// ---- POUs/Tc3 Objects/Alarm/GVL_FB_Alarm_1.TcGVL
{attribute 'Tc2GvlVarNames'}
VAR_GLOBAL CONSTANT
	nALARM_MAX_NO			:INT := 63;			(* Maximal number of alarms *)
END_VAR

// ---- POUs/Tc3 Objects/Communication/TCPIP/GVL_TCPIP.TcGVL
{attribute 'qualified_only'}
VAR_GLOBAL CONSTANT
	BUFFER_SIZE						:UDINT := 1000;(* Max. internal fifo/receiver buffer size *)

	CLIENT_SEND_CYCLE_TIME			:TIME := T#1S;
	RECEIVE_POLLING_TIME			:TIME := T#100MS;
	RECEIVE_MESSAGE_MAX				:UINT := 10;

	(* Some project specific error codes *)
	ERROR_RECEIVE_TIMEOUT			:UDINT := 16#8101;(* Receive timeout *)
	ERROR_SENDFIFO_OVERFLOW			:UDINT := 16#8102;(* Send fifo overflow *)
	ERROR_RECFIFO_OVERFLOW			:UDINT := 16#8103;(* Receive fifo overflow *)
END_VAR

// ---- POUs/Tc3 Objects/ExternalHardware/Gefran/GVL_GFX4IR.TcGVL
{attribute 'qualified_only'}
VAR_GLOBAL CONSTANT
	nZONES_MAX_NO			:UINT := 4;			(* Amount of control zones *)
END_VAR

// ---- POUs/Tc3 Objects/File/CSV/GVL_CSV.TcGVL
VAR_GLOBAL CONSTANT
	MAX_CSV_ROWS 					:UDINT := 50;
	MAX_CSV_COLUMNS 				:UDINT := 50;
	MAX_CSV_FIELD_LENGTH			:UDINT := 100;
END_VAR

// ---- POUs/Tc3 Objects/File/TXT/GVL_FB_LoadFromFile_1.TcGVL
{attribute 'Tc2GvlVarNames'}
VAR_GLOBAL CONSTANT
	usnFileArrayMaxDimR					:USINT := 100;		(* 0..usnMaxDimR - Number of rows to read. *)
	usnFileArrayMaxDimC					:USINT := 4;  		(* 0..usnMaxDimC -  Number of columns to read. *)
END_VAR

// ---- POUs/Tc3 Objects/Logger/GVL_Logger.TcGVL
{attribute 'Tc2GvlVarNames'}
VAR_GLOBAL
	unLOG_INSTANCE_IDX				:UINT;
END_VAR
VAR_GLOBAL CONSTANT
	sLOG_FILE_PATH					:STRING := '\Hard Disk\Riex\Log\';			(* Login file path *)
	sLOG_FILE_SUFFIX					:STRING := 'log';							(* Suffix of loggin file *)
	unNUM_OF_LOG_VAR					:UINT := 4;								(* Number of logging variables *)
	unLOG_MAX_NO						:UINT := 1;
	unLOG_BEFOR_MAX_NO				:UINT := 10;
	unLOG_DURING_MAX_NO				:UINT := 250;
	unLOG_AFTER_MAX_NO				:UINT := 10;
END_VAR

// ---- POUs/Tc3 Objects/Traceability/GVL_Trace.TcGVL
{attribute 'Tc2GvlVarNames'}
VAR_GLOBAL CONSTANT
	MAX_TRACE_ROWS 					:UDINT := 1;
	MAX_TRACE_COLUMNS 				:UDINT := 30;
	MAX_TRACE_FIELD_LENGTH			:UDINT := 100;
END_VAR

// ---- POUs/MAIN.TcPOU
PROGRAM MAIN
VAR
	tonDelay			:TON;

	lrRight:LREAL;
	lrRight2:WORD;
	lrClamp2Pos:LREAL;
	lrActSawingAngle :LREAL;
END_VAR


Init();										(* Call Init *)
tonDelay(IN := TRUE, PT := t#3s);
Gr00Coordinator(bEnable := tonDelay.Q);			(* Call Program *)
Gr01Coordinator(bEnable := tonDelay.Q);			(* Call Program *)
Gr05Coordinator(bEnable := tonDelay.Q);			(* Call Program *)


lrActSawingAngle := (45 / 180 * PI);

lrClamp2Pos := F_AxisClamp2Pos(
					bEnable := TRUE,
					lrActClamp2Pos := Gr05Control.fbCylinderPos.lrActPosition,
					lrAngle := lrActSawingAngle,
					lrRadius := stgGr01HMI.stHMITOPLC.rPipeDiameter / 2.0,
					lrPipeClampWidth := lrgGr05PipeClampWidth,
					lrSawbandGuideWidth := lrgGr05SawbandGuideWidth
				);

lrRight := F_GetCylinderPos(		F_SetCylinderPos(SEL(stgGr05HMI.stHMITOPLC.bCylinderPosActive, Gr05Control.fbCylinderPos.lrActPosition, lrClamp2Pos),
																		lrgGr05CylinderPosOffset,
																		lrgGr05CylinderPosOriginShiftPos,
																		etgGr05CylinderPosDirection,
																		usngGr05CylinderPosCodingType),
														lrgGr05CylinderPosOffset,
														lrgGr05CylinderPosOriginShiftPos,
														etgGr05CylinderPosDirection,
														usngGr05CylinderPosCodingType)
									    + lrgGr05Clamp2Width ;



lrRight2 := F_SetCylinderPos(SEL(stgGr05HMI.stHMITOPLC.bCylinderPosActive, Gr05Control.fbCylinderPos.lrActPosition, lrClamp2Pos),
																		lrgGr05CylinderPosOffset,
																		lrgGr05CylinderPosOriginShiftPos,
																		etgGr05CylinderPosDirection,
																		usngGr05CylinderPosCodingType);

END_PROGRAM

// ---- POUs/Init.TcPOU
PROGRAM Init
VAR
	bFirstTime					:BOOL; 				(* False = first run / True = not first run *)
END_VAR
VAR PERSISTENT
	bFirstTimePersistent			:BOOL;				(* Persistente Daten initialisieren *)
END_VAR


IF NOT bFirstTime
THEN
	A_InitGr0000();
	A_InitGr0100();
	A_InitGr0200();
	A_InitGr0500();

	bFirstTime:= TRUE;
END_IF

IF NOT bFirstTimePersistent
THEN

	bFirstTimePersistent:= TRUE;
END_IF

ACTION A_InitGr0000:
;
END_ACTION

ACTION A_InitGr0100:
;
END_ACTION

ACTION A_InitGr0200:
;
END_ACTION

ACTION A_InitGr0500:
;
END_ACTION

END_PROGRAM

// ---- POUs/Machine/Group_0000 - General/Gr00Coordinator.TcPOU
PROGRAM Gr00Coordinator
VAR_INPUT
	(* Input variables / Eingang Variablen *)
	bEnable					:BOOL;						(* Enable Group00 *)
END_VAR
VAR
	(* Enummerations *)

	(* Variables *)

	(* References *)

	(* Interfaces *)

	(* Instances *)

END_VAR

IF NOT bEnable
THEN
	RETURN;
END_IF;

Gr00Persistent(bEnable := TRUE);			(* Call Program *)
Gr00Simulation(bEnable := TRUE);			(* Call Program *)
Gr00MachineMode(bEnable := TRUE);		(* Call Program *)
Gr00Control(bEnable := TRUE);				(* Call Program *)
Gr00HMI(bEnable := TRUE);				(* Call Program *)

END_PROGRAM

// ---- POUs/Machine/Group_0000 - General/Gr00Persistent/Gr00Persistent.TcPOU
PROGRAM Gr00Persistent
VAR_INPUT
	(* Input variables / Eingang Variablen *)
	bEnable					:BOOL;						(* Enable Gr00Persistent *)
END_VAR
VAR PERSISTENT
	(* Enummerations *)

	(* Variables *)
	rOverride							:REAL;						(* Override 0 - 100 % *)
	udnCounterTotal						:UDINT;						(* Total counter *)
	udnCounterUser						:UDINT;						(* User counter *)
	bProgramActive						:BOOL;						(* Program active *)

	arstSaveDiagSlaveInfo 				:ARRAY [0..dnDIAG_SLAVEINFO_SIZE] OF ST_SlaveStateInfo;
	arstSaveDiagSlaveInfoScanned			:ARRAY [0..dnDIAG_SLAVEINFO_SIZE] OF ST_SlaveStateInfoScanned;

	(* References *)

	(* Interfaces *)

	(* Instances *)
END_VAR
VAR
	(* Enummerations *)

	(* Variables *)
	bFirstTime							:BOOL;

	(* References *)

	(* Interfaces *)

	(* Instances *)

END_VAR

IF NOT bEnable
THEN
	bFirstTime := FALSE;
	RETURN;
END_IF;

IF NOT bFirstTime
THEN
	A_SetPerVar();

	bFirstTime := TRUE;
END_IF;

A_GetPerVar();

ACTION A_GetPerVar:

bgGr00WritePersistent := rOverride <> stgGr00HMI.stHMITOPLC.rOverride
					OR udnCounterTotal <> stgGr00HMI.stPLCTOHMI.udnCounterTotal
					OR udnCounterUser <> stgGr00HMI.stPLCTOHMI.udnCounterUser
					OR bProgramActive <> stgGr00HMI.stHMITOPLC.bProgramActive
					OR MEMCMP(ADR(arstSaveDiagSlaveInfo), ADR(SaveDiagSlaveInfo), SIZEOF(SaveDiagSlaveInfo)) <> 0
					OR MEMCMP(ADR(arstSaveDiagSlaveInfoScanned), ADR(SaveDiagSlaveInfoScanned), SIZEOF(SaveDiagSlaveInfoScanned)) <> 0;

rOverride := stgGr00HMI.stHMITOPLC.rOverride;
udnCounterTotal := stgGr00HMI.stPLCTOHMI.udnCounterTotal;
udnCounterUser := stgGr00HMI.stPLCTOHMI.udnCounterUser;
bProgramActive := stgGr00HMI.stHMITOPLC.bProgramActive;

MEMCPY(ADR(arstSaveDiagSlaveInfo), ADR(SaveDiagSlaveInfo), SIZEOF(SaveDiagSlaveInfo));
MEMCPY(ADR(arstSaveDiagSlaveInfoScanned), ADR(SaveDiagSlaveInfoScanned), SIZEOF(SaveDiagSlaveInfoScanned));
END_ACTION

ACTION A_SetPerVar:

stgGr00HMI.stHMITOPLC.rOverride := rOverride;
stgGr00HMI.stPLCTOHMI.udnCounterTotal := udnCounterTotal;
stgGr00HMI.stPLCTOHMI.udnCounterUser := udnCounterUser;
stgGr00HMI.stHMITOPLC.bProgramActive := bProgramActive;

MEMCPY(ADR(SaveDiagSlaveInfo), ADR(arstSaveDiagSlaveInfo), SIZEOF(arstSaveDiagSlaveInfo));
MEMCPY(ADR(SaveDiagSlaveInfoScanned), ADR(arstSaveDiagSlaveInfoScanned), SIZEOF(arstSaveDiagSlaveInfoScanned));
END_ACTION

END_PROGRAM

// ---- POUs/Machine/Group_0000 - General/Gr00Simulation/Gr00Simulation.TcPOU
PROGRAM Gr00Simulation
VAR_INPUT
	(* Input variables / Eingang Variablen *)
	bEnable								:BOOL;						(* Enable Gr05Persistent *)
END_VAR
VAR
	(* Enummerations *)

	(* Variables *)

	(* References *)

	(* Interfaces *)

	(* Instances *)

END_VAR

IF NOT bEnable
THEN

	RETURN;
END_IF;

A_ForceInput();

ACTION A_ForceInput:


GVL_Gr00IO.binGr00AirPressureOK := TRUE;
GVL_Gr00IO.binGr00LightCurtainOK := TRUE;
GVL_Gr00IO.arbinGr00PowerSupplyOn[2] := TRUE;
GVL_Gr00IO.arbinGr00PowerSupplyOn[3] := TRUE;
GVL_Gr00IO.arbinGr00PowerSupplyOn[4] := TRUE;
GVL_Gr00IO.arbinGr00PowerSupplyOn[5] := TRUE;
GVL_Gr00IO.arbinGr00DoorsClosed[1] := TRUE;
GVL_Gr00IO.arbinGr00DoorsClosed[2] := TRUE;
GVL_Gr00IO.arbinGr00DoorsClosed[3] := TRUE;
GVL_Gr00IO.arbinGr00DoorsClosed[4] := TRUE;
GVL_Gr00IO.arbinGr00DoorsClosed[5] := TRUE;
GVL_Gr00IO.binGr00AllDoorsClosed := GVL_Gr00IO.arbinGr00DoorsClosed[1]
								AND GVL_Gr00IO.arbinGr00DoorsClosed[2]
								AND GVL_Gr00IO.arbinGr00DoorsClosed[3]
								AND GVL_Gr00IO.arbinGr00DoorsClosed[4]
								AND GVL_Gr00IO.arbinGr00DoorsClosed[5];

GVL_Gr00IO.binGr00AllDoorsLocked := TRUE;
GVL_Gr00IO.binGr00TempOK := TRUE;


// only for simulation
// GVL_Gr00IO.binNoEmergencyStop := TRUE;
// GVL_Gr00IO.binMoveRelease := TRUE;
// GVL_Gr00IO.binMoveReleaseSB := TRUE;
END_ACTION

END_PROGRAM

// ---- POUs/Machine/Group_0000 - General/Gr00MachineMode/Gr00MachineMode.TcPOU
PROGRAM Gr00MachineMode
VAR_INPUT
	(* Input variables / Eingang Variablen *)
	bEnable					:BOOL;						(* Enable Gr00MachineMode *)
END_VAR
VAR
	(* Enummerations *)

	(* Variables *)

	(* References *)

	(* Interfaces *)

	(* Instances *)

END_VAR

IF NOT bEnable
THEN
	RETURN;
END_IF;

Gr00Auto(bEnable := TRUE);			(* Call Program *)
Gr00Home(bEnable := TRUE);			(* Call Program *)
Gr00Manual(bEnable := TRUE);			(* Call Program *)

END_PROGRAM

// ---- POUs/Machine/Group_0000 - General/Gr00MachineMode/Gr00Auto/Gr00Auto.TcPOU
PROGRAM Gr00Auto
VAR_INPUT
	(* Input variables / Eingang Variablen *)
	bEnable					:BOOL;						(* Enable Gr00Auto *)
	bExecute				:BOOL;						(* Auto execute *)

	(* Instances *)
	fbInit						:FB_Gr00AutoInit;
	fbProcedure				:FB_Gr00AutoProcedure;
END_VAR
VAR
	(* Enummerations *)

	(* Variables *)

	(* References *)

	(* Interfaces *)

	(* Instances *)
	rtExecute					:R_TRIG;

	fbAlarm					:FB_Gr00AutoAlarm;
END_VAR
VAR CONSTANT
	nFatalErrorMaxIdx				:INT := 0;						(* Maximal index of  using alarms *)
	nErrorMaxIdx					:INT := 0;						(* Maximal index of  using alarms *)
	nWarningMaxIdx				:INT := 0;						(* Maximal index of  using alarms *)
	nMessageMaxIdx				:INT := 0;						(* Maximal index of  using alarms *)
	nHintMaxIdx					:INT := 0;						(* Maximal index of  using alarms *)

	dnFatalErrorBaseIdentNo		:DINT := 02000;				(* Fatal error identification number *)
	dnErrorBaseIdentNo			:DINT := 02100;				(* Error identification number *)
	dnWarningBaseIdentNo		:DINT := 02200;				(* Warning identification number *)
	dnMessageBaseIdentNo		:DINT := 02300;				(* Message identification number *)
	dnHintBaseIdentNo			:DINT := 02400;				(* Hint identification number *)
END_VAR

IF NOT bEnable
THEN
    RETURN;
END_IF;

(* Check auto execute *)
bExecute := bgGr00ModeAutomatic
		      AND NOT fbInit.bFirstTime;

rtExecute(CLK := bExecute);

IF rtExecute.Q
THEN
	A_Init();
END_IF;

A_Procedure();
A_Alarm();

ACTION A_Alarm:

(* Collect and execute input alarms *)
fbAlarm.stAlarmIn.arbError[0].bActive := FALSE;
fbAlarm.stAlarmIn.arbError[0].dnCode := dnErrorBaseIdentNo + 0;

fbAlarm(
	etMachineMode := etgGr00MachineMode,
	etMachineState := etgGr00MachineState,
	bNoEStop := bgGr00NoEmergencyStop,
	bConfirmAlarm := bgGr00ConfirmAlarm,
	dtDateTime := stgGr00DateTime.dtDateTime,
	nFatalErrorMaxIdx := nFatalErrorMaxIdx,
	nErrorMaxIdx := nErrorMaxIdx,
	nWarningMaxIdx := nWarningMaxIdx,
	nMessageMaxIdx := nMessageMaxIdx,
	nHintMaxIdx := nHintMaxIdx,
	bMoveInterrupted := bgGr00MoveInterrupted,
	bHomeCompleted := bgGr00HomeCompleted,
	stAlarmOut => stgGr00Alarm.stAuto
);
END_ACTION

ACTION A_Init:

(* Initializing variables *)
fbInit();
END_ACTION

ACTION A_Procedure:

(* Execute auto procedure *)
fbProcedure(
	bEnable := fbInit.bFirstTime,
	bExecute := etgGr00MachineState = ET_MachineState_eAutoExe
	             	       OR etgGr00MachineState = ET_MachineState_eAutoSteppingExe,
	bInterrupt := FALSE,
	bReleaseNextStep := etgGr00MachineState = ET_MachineState_eAutoExe
	             	       		       OR etgGr00MachineState = ET_MachineState_eAutoSteppingExe,
	bDone => bgGr00AutoCompleted,
	bInterrupted => bgGr00MoveInterrupted
);
END_ACTION

END_PROGRAM

// ---- POUs/Machine/Group_0000 - General/Gr00MachineMode/Gr00Home/Gr00Home.TcPOU
PROGRAM Gr00Home
VAR_INPUT
	(* Input variables / Eingang Variablen *)
	bEnable					:BOOL;						(* Enable Gr00Home *)
	bExecute				:BOOL;						(* Home execute *)

	(* Instances *)
	fbInit						:FB_Gr00HomeInit;
	fbProcedure				:FB_Gr00HomeProcedure;
END_VAR
VAR
	(* Enummerations *)

	(* Variables *)

	(* References *)

	(* Interfaces *)

	(* Instances *)
	rtExecute					:R_TRIG;

	fbAlarm					:FB_Gr00HomeAlarm;

END_VAR
VAR CONSTANT
	nFatalErrorMaxIdx				:INT := 0;						(* Maximal index of  using alarms *)
	nErrorMaxIdx					:INT := 0;						(* Maximal index of  using alarms *)
	nWarningMaxIdx				:INT := 0;						(* Maximal index of  using alarms *)
	nMessageMaxIdx				:INT := 0;						(* Maximal index of  using alarms *)
	nHintMaxIdx					:INT := 0;						(* Maximal index of  using alarms *)

	dnFatalErrorBaseIdentNo		:DINT := 03000;				(* Fatal error identification number *)
	dnErrorBaseIdentNo			:DINT := 03100;				(* Error identification number *)
	dnWarningBaseIdentNo		:DINT := 03200;				(* Warning identification number *)
	dnMessageBaseIdentNo		:DINT := 03300;				(* Message identification number *)
	dnHintBaseIdentNo			:DINT := 03400;				(* Hint identification number *)
END_VAR

IF NOT bEnable
THEN
	RETURN;
END_IF;

(* Check home execute *)
bExecute := etgGr00MachineState = ET_MachineState_eHomeRefExe
		      OR etgGr00MachineState = ET_MachineState_eHomeExe;

rtExecute(CLK := bExecute);                   

IF rtExecute.Q
THEN
	fbInit.bFirstTime := FALSE;
	A_Init();
END_IF;

A_Procedure();
A_Alarm();

ACTION A_Alarm:

(* Collect and execute input alarms *)
fbAlarm.stAlarmIn.arbError[0].bActive := fbProcedure.bErrorByProgramVerification;
fbAlarm.stAlarmIn.arbError[0].dnCode := dnErrorBaseIdentNo + 0;

fbAlarm(
	etMachineMode := etgGr00MachineMode,
	etMachineState := etgGr00MachineState,
	bNoEStop := bgGr00NoEmergencyStop,
	bConfirmAlarm := bgGr00ConfirmAlarm,
	dtDateTime := stgGr00DateTime.dtDateTime,
	nFatalErrorMaxIdx := nFatalErrorMaxIdx,
	nErrorMaxIdx := nErrorMaxIdx,
	nWarningMaxIdx := nWarningMaxIdx,
	nMessageMaxIdx := nMessageMaxIdx,
	nHintMaxIdx := nHintMaxIdx,
	bMoveInterrupted := bgGr00MoveInterrupted,
	bHomeCompleted := bgGr00HomeCompleted,
	stAlarmOut => stgGr00Alarm.stHome
);
END_ACTION

ACTION A_Init:

(* Initializing variables *)
fbInit();
END_ACTION

ACTION A_Procedure:

(* Execute home procedure *)
fbProcedure(
	bEnable := etgGr00MachineMode = ET_MachineMode_eHome,
	bExecute := rtExecute.Q,
	bReleaseNextStep := etgGr00MachineState = ET_MachineState_eHomeRefExe
		      	     		      OR etgGr00MachineState = ET_MachineState_eHomeExe
);
END_ACTION

END_PROGRAM

// ---- POUs/Machine/Group_0000 - General/Gr00MachineMode/Gr00Manual/Gr00Manual.TcPOU
PROGRAM Gr00Manual
VAR_INPUT
	(* Input variables / Eingang Variablen *)
	bEnable					:BOOL;						(* Enable Gr00Manual *)
	bExecute				:BOOL;						(* Manual execute *)

	(* Instances *)
	fbInit						:FB_Gr00ManualInit;
	fbProcedure				:FB_Gr00ManualProcedure;
END_VAR
VAR
	(* Enummerations *)

	(* Variables *)

	(* References *)

	(* Interfaces *)

	(* Instances *)
	rtExecute					:R_TRIG;

	fbAlarm					:FB_Gr00ManualAlarm;
END_VAR
VAR CONSTANT
	nFatalErrorMaxIdx				:INT := 0;						(* Maximal index of  using alarms *)
	nErrorMaxIdx					:INT := 0;						(* Maximal index of  using alarms *)
	nWarningMaxIdx				:INT := 0;						(* Maximal index of  using alarms *)
	nMessageMaxIdx				:INT := 0;						(* Maximal index of  using alarms *)
	nHintMaxIdx					:INT := 0;						(* Maximal index of  using alarms *)

	dnFatalErrorBaseIdentNo		:DINT := 04000;				(* Fatal error identification number *)
	dnErrorBaseIdentNo			:DINT := 04100;				(* Error identification number *)
	dnWarningBaseIdentNo		:DINT := 04200;				(* Warning identification number *)
	dnMessageBaseIdentNo		:DINT := 04300;				(* Message identification number *)
	dnHintBaseIdentNo			:DINT := 04400;				(* Hint identification number *)
END_VAR

IF NOT bEnable
THEN
	RETURN;
END_IF;

(* Check manual execute *)
bExecute := etgGr00MachineMode = ET_MachineMode_eManual;

rtExecute(CLK := bExecute);

IF rtExecute.Q
THEN
	fbInit.bFirstTime := FALSE;
	A_Init();
END_IF;

A_Procedure();
A_Alarm();

ACTION A_Alarm:

(* Collect and execute input alarms *)
fbAlarm.stAlarmIn.arbError[0].bActive := FALSE;
fbAlarm.stAlarmIn.arbError[0].dnCode := dnErrorBaseIdentNo + 0;

fbAlarm(
	etMachineMode := etgGr00MachineMode,
	etMachineState := etgGr00MachineState,
	bNoEStop := bgGr00NoEmergencyStop,
	bConfirmAlarm := bgGr00ConfirmAlarm,
	dtDateTime := stgGr00DateTime.dtDateTime,
	nFatalErrorMaxIdx := nFatalErrorMaxIdx,
	nErrorMaxIdx := nErrorMaxIdx,
	nWarningMaxIdx := nWarningMaxIdx,
	nMessageMaxIdx := nMessageMaxIdx,
	nHintMaxIdx := nHintMaxIdx,
	bHomeCompleted := bgGr00HomeCompleted,
	stAlarmOut => stgGr00Alarm.stManual
);
END_ACTION

ACTION A_Init:

(* Initializing variables *)
fbInit();
END_ACTION

ACTION A_Procedure:

(* Execute manual procedure *)
fbProcedure(
	bEnable := etgGr00MachineMode = ET_MachineMode_eManual,
	bExecute := rtExecute.Q,
	bReleaseNextStep := etgGr00MachineMode = ET_MachineMode_eManual
);
END_ACTION

END_PROGRAM

// ---- POUs/Machine/Group_0000 - General/Gr00Control/Gr00Control.TcPOU
PROGRAM Gr00Control
VAR_INPUT
	(* Input variables / Eingang Variablen *)
	bEnable					:BOOL;						(* Enable Gr00Control *)

	fbProgram				:FB_Gr00Program;
END_VAR
VAR
	(* Enummerations *)

	(* Variables *)

	(* References *)

	(* Interfaces *)

	(* Instances *)
	fbAlarm					:FB_Gr00Alarm;
	fbSafety					:FB_Gr00Safety;
	fbSignals				:FB_Gr00Signals;
	fbUtility					:FB_Gr00Utility;
	fbPeriphery				:FB_Gr00Periphery;

	ftClampsChecked			:F_TRIG;
	tonClampsChecked		:TON;
	fbMachineStandstill		:FB_SignalHandlingDelay;

	fbStartHMI				:NT_StartProcess;
	tonStartHmi				:TON;

END_VAR
VAR CONSTANT
	nFatalErrorMaxIdx				:INT := 1;						(* Maximal index of  using alarms *)
	nErrorMaxIdx					:INT := 12;					(* Maximal index of  using alarms *)
	nWarningMaxIdx				:INT := 0;						(* Maximal index of  using alarms *)
	nMessageMaxIdx				:INT := 4;						(* Maximal index of  using alarms *)
	nHintMaxIdx					:INT := 0;						(* Maximal index of  using alarms *)

	dnFatalErrorBaseIdentNo		:DINT := 01000;				(* Fatal error identification number *)
	dnErrorBaseIdentNo			:DINT := 01100;				(* Error identification number *)
	dnWarningBaseIdentNo		:DINT := 01200;				(* Warning identification number *)
	dnMessageBaseIdentNo		:DINT := 01300;				(* Message identification number *)
	dnHintBaseIdentNo			:DINT := 01400;				(* Hint identification number *)
END_VAR

IF NOT bEnable
THEN
	RETURN;
END_IF;

A_Periphery();
A_Utility();
A_Program();
A_Safety();
A_Signals();
A_Alarm();
A_HMI();

ACTION A_Alarm:

(* Collect and execute input alarms *)
fbAlarm.stAlarmIn.arbFatalError[0].bActive := fbSafety.fbNoEmergencyStop.bError;
fbAlarm.stAlarmIn.arbFatalError[0].dnCode := dnFatalErrorBaseIdentNo + 0;

fbAlarm.stAlarmIn.arbError[0].bActive := NOT binGr00LightCurtainOK
                                                		      AND (Gr01Home.fbProcedure.bBusy
                                                      				OR Gr01Auto.fbProcedure.bBusy);
fbAlarm.stAlarmIn.arbError[0].dnCode := dnErrorBaseIdentNo + 0;

fbAlarm.stAlarmIn.arbError[1].bActive := fbSafety.fbAirPressure.bError;
fbAlarm.stAlarmIn.arbError[1].dnCode := dnErrorBaseIdentNo + 1;

fbAlarm.stAlarmIn.arbError[2].bActive := FALSE;
fbAlarm.stAlarmIn.arbError[2].dnCode := dnErrorBaseIdentNo + 2;

fbAlarm.stAlarmIn.arbError[4].bActive := NOT fbSafety.bFieldbusMasterOK AND fbSafety.fbFieldbus.bInit;
fbAlarm.stAlarmIn.arbError[4].dnCode := dnErrorBaseIdentNo + 4;

fbAlarm.stAlarmIn.arbError[5].bActive := fbSafety.bFieldbusBrake;
fbAlarm.stAlarmIn.arbError[5].dnCode := dnErrorBaseIdentNo + 5;

fbAlarm.stAlarmIn.arbError[6].bActive := fbSafety.fbTemperatur.bError;
fbAlarm.stAlarmIn.arbError[6].dnCode := dnErrorBaseIdentNo + 6;

fbAlarm.stAlarmIn.arbError[7].bActive := NOT fbSafety.arbPowerSupplyOn[1];
fbAlarm.stAlarmIn.arbError[7].dnCode := dnErrorBaseIdentNo + 7;

fbAlarm.stAlarmIn.arbError[8].bActive :=NOT fbSafety.arbPowerSupplyOn[2];
fbAlarm.stAlarmIn.arbError[8].dnCode := dnErrorBaseIdentNo + 8;

fbAlarm.stAlarmIn.arbError[9].bActive := NOT fbSafety.arbPowerSupplyOn[3];
fbAlarm.stAlarmIn.arbError[9].dnCode := dnErrorBaseIdentNo + 9;

fbAlarm.stAlarmIn.arbError[10].bActive := FALSE(*SystemInfo.bootDataFlags.5*);
fbAlarm.stAlarmIn.arbError[10].dnCode := dnErrorBaseIdentNo + 10;

fbAlarm.stAlarmIn.arbError[11].bActive := fbProgram.fbRead.bError
								      AND  fbProgram.fbRead.udnErrorNo <> 31;
fbAlarm.stAlarmIn.arbError[11].dnCode := dnErrorBaseIdentNo + 11;

fbAlarm.stAlarmIn.arbError[12].bActive := fbProgram.fbRead.bError
								      AND  fbProgram.fbRead.udnErrorNo = 31;
fbAlarm.stAlarmIn.arbError[12].dnCode := dnErrorBaseIdentNo + 12;

fbAlarm.stAlarmIn.arbWarning[0].bActive := fbSafety.fbTemperatur.bWarning;
fbAlarm.stAlarmIn.arbWarning[0].dnCode := dnWarningBaseIdentNo + 0;

fbAlarm.stAlarmIn.arbWarning[1].bActive := NOT GVL_Gr00IO.binGr00Luetze_F1;
fbAlarm.stAlarmIn.arbWarning[1].dnCode := dnWarningBaseIdentNo + 1;

fbAlarm.stAlarmIn.arbWarning[2].bActive := NOT GVL_Gr00IO.binGr00Luetze_F2;
fbAlarm.stAlarmIn.arbWarning[2].dnCode := dnWarningBaseIdentNo + 2;

fbAlarm.stAlarmIn.arbWarning[3].bActive := NOT GVL_Gr00IO.binGr00Luetze_F3;
fbAlarm.stAlarmIn.arbWarning[3].dnCode := dnWarningBaseIdentNo + 3;

fbAlarm.stAlarmIn.arbWarning[4].bActive := NOT GVL_Gr00IO.binGr00PS6A24Warning_1;
fbAlarm.stAlarmIn.arbWarning[4].dnCode := dnWarningBaseIdentNo + 4;

fbAlarm.stAlarmIn.arbWarning[5].bActive := NOT GVL_Gr00IO.binGr00PS6A24Warning_2;
fbAlarm.stAlarmIn.arbWarning[5].dnCode := dnWarningBaseIdentNo + 5;

fbAlarm.stAlarmIn.arbWarning[6].bActive := NOT GVL_Gr00IO.binGr00PS6A24Ready;
fbAlarm.stAlarmIn.arbWarning[6].dnCode := dnWarningBaseIdentNo + 6;

fbAlarm.stAlarmIn.arbMessage[0].bActive := fbSafety.fbAirPressure.udnMessageNo = 1;
fbAlarm.stAlarmIn.arbMessage[0].dnCode := dnMessageBaseIdentNo + 0;

fbAlarm.stAlarmIn.arbMessage[1].bActive := stgGr00HMI.stHMITOPLC.bSafetyInterlockOff;
fbAlarm.stAlarmIn.arbMessage[1].dnCode := dnMessageBaseIdentNo + 1;

fbAlarm.stAlarmIn.arbMessage[2].bActive := NOT binGr00LightCurtainOK
                                            				      AND NOT fbAlarm.stAlarmIn.arbError[0].bActive
                                            				      AND NOT stgGr00Alarm.stControl.arbError[0].bActive;
fbAlarm.stAlarmIn.arbMessage[2].dnCode := dnMessageBaseIdentNo + 2;

fbAlarm.stAlarmIn.arbMessage[4].bActive := NOT binGr00AllDoorsClosed;
fbAlarm.stAlarmIn.arbMessage[4].dnCode := dnMessageBaseIdentNo + 4;

(* Execute utility *)
fbAlarm(
	etMachineMode := etgGr00MachineMode,
	etMachineState := etgGr00MachineState,
	bNoEStop := bgGr00NoEmergencyStop,
	bConfirmAlarm := bgGr00ConfirmAlarm,
	dtDateTime := stgGr00DateTime.dtDateTime,
	nFatalErrorMaxIdx := nFatalErrorMaxIdx,
	nErrorMaxIdx := nErrorMaxIdx,
	nWarningMaxIdx := nWarningMaxIdx,
	nMessageMaxIdx := nMessageMaxIdx,
	nHintMaxIdx := nHintMaxIdx,
	bMoveInterrupted := bgGr00MoveInterrupted,
	bHomeCompleted := bgGr00HomeCompleted,
	stAlarmOut => stgGr00Alarm.stControl
);
END_ACTION

ACTION A_HMI:
(*Starting the HMI*)

tonStartHmi(IN:=TRUE, PT:= T#2s);

fbStartHMI(
		PATHSTR   := 'C:\Riex\HMI\App.exe',
    		DIRNAME   :='C:\Riex\HMI\',
    		START     := tonStartHmi.Q,
		TMOUT     := T#5s
		);
END_ACTION

ACTION A_Periphery:

(* Periphery *)
fbPeriphery(
	bEnable := TRUE,
	Periphery := Periphery
);
END_ACTION

ACTION A_Program:

(* Execute program *)
fbProgram(
	sPath := sgGr00PrgPath,
	sName := sgGr00PrgName,
	sSuffix := sgGr00PrgSuffix
);
END_ACTION

ACTION A_Safety:

bgGr00DoorsUnlockRelease := bgGr00ModeManual
						        OR
							(bgGr00ModeHome
							 AND NOT bgGr00MachineRunning)
						        OR
							(bgGr00ModeAutomatic
							 AND NOT bgGr00MachineRunning);

(* Execute safety *)
fbSafety(
	etMachineMode := etgGr00MachineMode,
	etMachineState := etgGr00MachineState,
	bNoEStop := binGr00NoEmergencyStop,
	bConfirmEStop := FALSE,
	bMachineRunning := bgGr00MachineRunning,
	arbPowerSupplyOn := arbinGr00PowerSupplyOn,
	bLightCurtain := binGr00LightCurtainOK,
	bConfirmLightCurtain := (bgGr00ConfirmAlarm
						OR etgGr00MachineMode = ET_MachineMode_eManual
						OR etgGr00MachineMode = ET_MachineMode_eHome
						OR etgGr00MachineMode = ET_MachineMode_eAutomatic
						OR stgGr00HMI.stHMITOPLC.bSafetyInterlockOff)
						AND NOT stgGr00Alarm.stControl.arbError[0].bActive,
	bAirPressure := binGr00AirPressureOK,
	arbDoorsClosed := arbinGr00DoorsClosed,
	bDoorsClosed := binGr00AllDoorsClosed,
	bDoorsLocked := binGr00AllDoorsLocked,
	bTemperatur := binGr00TempOK,
	stFieldbusStatus := stinGr00FieldbusStatus,
	tFieldbusMasterStartUp := tgGr00FieldbusMasterStartUp,
	tPowerSupplyOn := tgGr00PowerSupplyOn,
	tPowerSupplyOff := tgGr00PowerSupplyOff,
	tAirPressureOnDelay := tgGr00AirPressureOnDelay,
	tAirPresentDelay := tgGr00AirPressureDelay,
	tAirPressureBuildUp := tgGr00AirPressureBuildUp,
	tLightCurtainDelay := tgGr00LightCurtainDelay,
	tAdsTimeOut := DEFAULT_ADS_TIMEOUT,
	bNoEmergencyStop => bgGr00NoEmergencyStop,
	bAirPressureOK => bgGr00AirPressureOK,
	bAirPressureOn => boutGr00AirPressureOn,
	bPowerSupplyOk => bgGr00PowerSupplyOk,
	bLightCurtainOK => bgGr00LightCurtainOK,
	bConfirmedLightCurtain => boutGr00ConfLightCurtain,
	bAllDoorsLock => boutGr00AllDoorsLock,
	bAllDoorsClosed => bgGr00AllDoorsClosed,
	bAllDoorsClosedLocked => bgGr00AllDoorsClosedLocked
);
END_ACTION

ACTION A_Signals:

(* Collect and execute input signals *)
fbSignals.stAlarm.bFatalError := stgGr00Alarm.stControl.bFatalError OR stgGr00Alarm.stManual.bFatalError OR stgGr00Alarm.stHome.bFatalError OR stgGr00Alarm.stAuto.bFatalError
							OR stgGr01Alarm.stControl.bFatalError OR stgGr01Alarm.stManual.bFatalError OR stgGr01Alarm.stHome.bFatalError OR stgGr01Alarm.stAuto.bFatalError
							OR stgGr02Alarm.stControl.bFatalError OR stgGr02Alarm.stManual.bFatalError OR stgGr02Alarm.stHome.bFatalError OR stgGr02Alarm.stAuto.bFatalError
							OR stgGr05Alarm.stControl.bFatalError OR stgGr05Alarm.stManual.bFatalError OR stgGr05Alarm.stHome.bFatalError OR stgGr05Alarm.stAuto.bFatalError;
fbSignals.stAlarm.bError := stgGr00Alarm.stControl.bError OR stgGr00Alarm.stManual.bError OR stgGr00Alarm.stHome.bError OR stgGr00Alarm.stAuto.bError
						OR stgGr01Alarm.stControl.bError OR stgGr01Alarm.stManual.bError OR stgGr01Alarm.stHome.bError OR stgGr01Alarm.stAuto.bError
						OR stgGr02Alarm.stControl.bError OR stgGr02Alarm.stManual.bError OR stgGr02Alarm.stHome.bError OR stgGr02Alarm.stAuto.bError
						OR stgGr05Alarm.stControl.bError OR stgGr05Alarm.stManual.bError OR stgGr05Alarm.stHome.bError OR stgGr05Alarm.stAuto.bError;
fbSignals.stAlarm.bWarning := stgGr00Alarm.stControl.bWarning OR stgGr00Alarm.stManual.bWarning OR stgGr00Alarm.stHome.bWarning OR stgGr00Alarm.stAuto.bWarning
		        					OR stgGr01Alarm.stControl.bWarning OR stgGr01Alarm.stManual.bWarning OR stgGr01Alarm.stHome.bWarning OR stgGr01Alarm.stAuto.bWarning
		        					OR stgGr02Alarm.stControl.bWarning OR stgGr02Alarm.stManual.bWarning OR stgGr02Alarm.stHome.bWarning OR stgGr02Alarm.stAuto.bWarning
		        					OR stgGr05Alarm.stControl.bWarning OR stgGr05Alarm.stManual.bWarning OR stgGr05Alarm.stHome.bWarning OR stgGr05Alarm.stAuto.bWarning;
fbSignals.stAlarm.bMessage := stgGr00Alarm.stControl.bMessage OR stgGr00Alarm.stManual.bMessage OR stgGr00Alarm.stHome.bMessage OR stgGr00Alarm.stAuto.bMessage
		        					OR stgGr01Alarm.stControl.bMessage OR stgGr01Alarm.stManual.bMessage OR stgGr01Alarm.stHome.bMessage OR stgGr01Alarm.stAuto.bMessage
		        					OR stgGr02Alarm.stControl.bMessage OR stgGr02Alarm.stManual.bMessage OR stgGr02Alarm.stHome.bMessage OR stgGr02Alarm.stAuto.bMessage
		        					OR stgGr05Alarm.stControl.bMessage OR stgGr05Alarm.stManual.bMessage OR stgGr05Alarm.stHome.bMessage OR stgGr05Alarm.stAuto.bMessage;
fbSignals.stAlarm.bHint := stgGr00Alarm.stControl.bHint OR stgGr00Alarm.stManual.bHint OR stgGr00Alarm.stHome.bHint OR stgGr00Alarm.stAuto.bHint
	       					OR stgGr01Alarm.stControl.bHint OR stgGr01Alarm.stManual.bHint OR stgGr01Alarm.stHome.bHint OR stgGr01Alarm.stAuto.bHint
	       					OR stgGr02Alarm.stControl.bHint OR stgGr02Alarm.stManual.bHint OR stgGr02Alarm.stHome.bHint OR stgGr02Alarm.stAuto.bHint
	       					OR stgGr05Alarm.stControl.bHint OR stgGr05Alarm.stManual.bHint OR stgGr05Alarm.stHome.bHint OR stgGr05Alarm.stAuto.bHint;

(* Execute signals *)
fbSignals(
	etMachineMode := etgGr00MachineMode,
	etMachineState := etgGr00MachineState,
	bMachineRunning := bgGr00MachineRunning,
	stBlinker => stgGr00Blinker,
	bBulbBtnStart => boutGr00BulbBtnStart,
	bBulbBtnStop => boutGr00BulbBtnStop,
	bBulbBtnHome => boutGr00BulbBtnHome,
	bBulbGreen => boutGr00BulbGreen,
	bBulbRed => boutGr00BulbRed,
	bBulbYellow => boutGr00BulbYellow,
	bHorn => boutGr00Horn
);

(* Signal button bulb "reset" / Signallampe "Reset" *)
boutGr00BulbBtnReset := binGr00NoEmergencyStop OR stgGr00Blinker.Q1;
END_ACTION

ACTION A_Utility:

(* Execute utility *)
fbUtility(
	bSignalStart := binGr00PushBtnStart OR stgGr00HMI.stHMITOPLC.bBtnStart,
	bSignalStop :=NOT binGr00PushBtnStop OR stgGr00HMI.stHMITOPLC.bBtnStop,
	bSignalAbort := fbSignals.stAlarm.bFatalError
				     OR fbSignals.stAlarm.bError,
	bSignalHome := binGr00PushBtnHome,
	bSignalReference := binGr00PushBtnRef OR stgGr00HMI.stHMITOPLC.bBtnForceRef,
	bSignalReset := binGr00PushBtnReset OR stgGr00HMI.stHMITOPLC.bBtnReset,
	bSignalMachinePurge := stgGr00HMI.stHMITOPLC.bBtnMachinePurge,
	bAutoStartRelease := binGr01SawbandRelease
					       AND bgGr05PipeEndPresent
					       AND (stgGr05HMI.stHMITOPLC.bCylinderPosActive
							  OR stgGr05HMI.stPLCTOHMI.arlrAxisClampActPos[2] < ABS(99999.0))
					       AND NOT stgGr05Alarm.stAuto.arbWarning[0].bActive,
	bHomeStartRelease := (stgGr05HMI.stHMITOPLC.bCylinderPosActive
							  OR stgGr05HMI.stPLCTOHMI.arlrAxisClampActPos[2] < ABS(99999.0)),
	bAutoToHome := NOT stgGr05Alarm.stAuto.arbWarning[0].bActive,
	bHomeCompleted := bgGr00HomeCompleted
					     AND bgGr01HomeCompleted
					     AND bgGr02HomeCompleted
					     AND bgGr05HomeCompleted,
	bAutoCompleted := bgGr00AutoCompleted
					  AND bgGr01AutoCompleted
					  AND bgGr02AutoCompleted
					  AND bgGr05AutoCompleted,
	bAllDoorsClosed := binGr00AllDoorsClosed,
	bAllDoorsLocked := bgGr00AllDoorsClosedLocked,
	bLightCurtainOk := bgGr00LightCurtainOK,
	etMachineModeReq := stgGr00HMI.stHMITOPLC.etMachineMode,
	bExeCounter := bgGr00AutoCompleted
					  AND bgGr01AutoCompleted
					  AND bgGr02AutoCompleted
					  AND bgGr05AutoCompleted,
	bResetCounterUser := stgGr00HMI.stHMITOPLC.bResetCounterUser,
	bStartTime := Gr01Control.fbUtility.arbStartProcess[1]
				OR Gr01Control.fbUtility.arbStartProcess[2]
				OR Gr01Control.fbUtility.arbStartProcess[3],
	bStopTime := bgGr01AutoCompleted
				OR Gr01Control.fbUtility.arbStopProcess[1]
				OR Gr01Control.fbUtility.arbStopProcess[2]
				OR Gr01Control.fbUtility.arbStopProcess[3],
	bLifetimeOn := TRUE,
	bResetLifetimeAll := FALSE,
	sLifetimeFilePath := sgGr00MachineLifetimeFilePath,
	sLifetimeFileName := sgGr00MachineLifetimeFileName,
	bWritePersistent :=  bgGr00WritePersistent
					  OR  bgGr01WritePersistent
					  OR  bgGr02WritePersistent
					  OR  bgGr05WritePersistent,
	bDownTraceDataExe := FALSE,
	rGlobalOverride := stgGr00HMI.stHMITOPLC.rOverride,
	udnCounterTotal := stgGr00HMI.stPLCTOHMI.udnCounterTotal,
	udnCounterUser := stgGr00HMI.stPLCTOHMI.udnCounterUser,
	tAdsTimeOut := DEFAULT_ADS_TIMEOUT,
	etMachineMode => etgGr00MachineMode,
	etMachineState => etgGr00MachineState,
	bModeAutomatic => bgGr00ModeAutomatic,
	bModeHome => bgGr00ModeHome,
	bModeManual => bgGr00ModeManual,
	bMachineRunning => bgGr00MachineRunning,
	bMachineStandstill => bgGr00MachineStandstill,
	bMachinePurge => bgGr00MachinePurge,
	bConfirmAlarm => bgGr00ConfirmAlarm,
	rActOverride => rgGr00Override,
	lrLifetimeAll => stgGr00HMI.stPLCTOHMI.lrMachineLifetime,
	lrLifetimeAfterTrunOn => stgGr00HMI.stPLCTOHMI.lrMachineLifetimeAfterTurnOn,
	lrActCycleTime => lrgActCycleTime,
	dwCycleTime => stgGr00HMI.stPLCTOHMI.dwCycleTime
);
END_ACTION

END_PROGRAM

// ---- POUs/Machine/Group_0000 - General/Gr00Control/Gr00Program/FB_Gr00Program.TcPOU
FUNCTION_BLOCK FB_Gr00Program
(*

The function block used to control general utility of the machine.

Constructor: 		Patryk Panylo
Company:		E. Riexinger GmbH
Date:			28.04.2015
Version:			1.00

Date:			Revision:		Who:				Comment
dd.mm.yyyy		x.xx			Initials			comment

*)
VAR_INPUT
	(* Input variables / Eingang Variablen *)
	bRead				:BOOL;						(* Read process parameters from file *)
	sPath				:STRING;					(* Program path e.g. '\Hard Disk\Riex\Recipe\'*)
	sName				:STRING;					(* Program name e.g. 'default' *)
	sSuffix				:STRING;					(* Program suffix e.g. 'prg' *)
END_VAR
VAR_OUTPUT
	(* Output variables / Ausgang Variablen *)

END_VAR
VAR_IN_OUT
	(* Input Output variables / Ausgang Variablen *)

END_VAR
VAR
	(* Enummerations *)

	(* Variables *)

	(* References *)

	(* Interfaces *)

	(* Instances *)
	fbRead				:FB_LoadFromFile;			(* Load program *)
END_VAR


A_Program();

ACTION A_Program:

fbRead(
	bEnable := TRUE,
	bExecute := bRead,
	byConfig := 4,
	sFilePath := sPath,
	sFileName := sName,
	sFileSuffix := sSuffix,
	sSep := ';',
	sEndLine:= '$N',
	sComment := '*',
	tTimeout := t#500ms
);

stgGr00HMI.stPLCTOHMI.sPrgFilePath := fbRead.sPathName;
END_ACTION

END_FUNCTION_BLOCK

// ---- POUs/Tc2 Objects/File/FB_LoadFromFile.TcPOU
FUNCTION_BLOCK FB_LoadFromFile
(*
Function to make easier work with file. Below options to choose. 
Chose option doasn't work with the others option. Allways is checking  only exist of file.
 
00000000 - 0 - Only check exist of file.
00000001 - 1 - Read line by line and save to array of string.
00000010 - 2 - Read line by line. Save first signs to string and convert to array of bool.
00000011 - 3 - Transfer  array form file to array of string on PLC - requirements:
			- kind of columns separator (bySep) and sign end of line (byEndLine),
			- amount of rows (usiMaxDimR) and columns (usiMaxDimR) to read.
00000111 - 4 - Option 3 + get real only real from string if capital letters then error

Constructor: 		Patryk Panylo
Company:		E. Riexinger GmbH
Date:			18.11.2015
Version:			1.00

Date:			Revision:		Who:				Comment
dd.mm.yyyy		x.xx			Initials			comment

*)
VAR_INPUT
	(* Enummerations *)

	(* Variables *)
	bEnable						:BOOL;									(* Enable FB *)
	bExecute					:BOOL; 									(* Execute load data *)
	byConfig 					:BYTE := 0;								(* Configuration byte
																		    Options:  - 2#00000000 (default),
																				    - 2#00000001 (actOption1),
																			  	    - 2#00000010 (actOption2),
																				    - 2#00000011 (actOption3),
																				    - 2#00000111 (actOption4),
																		*)
	sFilePath					:STRING;								(* File path *)
	sFileName					:STRING;								(* File name *)
	sFileSuffix					:STRING := 'dat';							(* Suffix of file *)
	sSep						:STRING := '$T'; 							(* Seperator sign for colums *)
	sEndLine					:STRING := '$N'; 							(* End line sign for lines *)
	sComment					:STRING := '!'; 							(* End line sign for lines *)
	tTimeout						:TIME := T#1s;							(* TimeOut *)

	(* References *)

	(* Interfaces *)


	(* Instances *)

END_VAR
VAR_OUTPUT
	(* Enummerations *)

	(* Variables *)
	arsData						:ARRAY [0..usnFileArrayMaxDimR] OF STRING [255];					(* Used with Option1 -  Array with read data from file in String[160] *)
	arbDataBool					:ARRAY [0..usnFileArrayMaxDimR] OF BOOL;							(* Used with Option2 - Array with read data from file in Bool *)
	arsDataDimRC				:ARRAY [0..usnFileArrayMaxDimR, 0..usnFileArrayMaxDimC ] OF STRING [20]; 		(* Used with Option3 - Matrix with read data from file in String[160] *)
	arrDataDimRC				:ARRAY [0..usnFileArrayMaxDimR, 0..usnFileArrayMaxDimC ] OF REAL; 			(* Matrix with read data from file in real *)
	bDone						:BOOL;													(* Program done *)
	bBusy						:BOOL;													(* Program busy *)
	bError						:BOOL;													(* Error *)
	udnErrorNo					:UDINT;													(* Error number *)
	sErrorMsg					:STRING; 												(* Error message *)

	(* References *)

	(* Interfaces *)

	(* Instances *)

END_VAR
VAR
	(* Enummerations *)
	etLoadFromFile				:ET_LoadFromFile;								(* Load from file enum variable *)

	(* Variables *)
	dwMode						:DWORD;										(* Contains the mode in which the file is to be opened *)
	sPathName					:STRING;										(* Contains the path and filename for the file to be opened *)
	hFileHandle					:UINT;											(* File handle *)
	usnRowsCounter				:USINT; 											(* Counter of rows (lines) in a  file*)

	sDataSign					:STRING[1];										(* Read first sign from line *)
	sDataString					:STRING[usnFileArrayMaxDimR];							(* Created string of sign *)
	arbyData					:ARRAY [0..usnFileArrayMaxDimR] OF BYTE;					(* String into array of byte *)
	ptString 						:POINTER TO ARRAY[0..usnFileArrayMaxDimR] OF BYTE;		(* Pointer to sDataString *)

	byDataSign					:BYTE;											(* Marker for sign form line *)
	ptByte						:POINTER TO BYTE;								(* Pointer to arsData *)
	usnColumnsCounter 			:USINT; 											(* Counter of colums *)

	bFirstTime					:BOOL;

	(* References *)

	(* Interfaces *)

	(* Instances *)
	tonTimeout					:TON;

	fbFileOpen					:FB_FileOpen;		(* Open file *)
	fbFileGets					:FB_FileGets;			(* Read from file *)
	fbFileClose					:FB_FileClose;		(* Close file *)

	rtExecute						:R_TRIG;				(* Positive edge for start *)

END_VAR

IF NOT bEnable
THEN
	bDone := FALSE;					(* Program done *)
	bBusy := FALSE;                                  	(* Program not busy *)
	bError := FALSE;                                 	(* Program not error *)
	udnErrorNo := 0;                                 		(* Error number *)

	bFirstTime := FALSE;
	RETURN;
END_IF;

IF NOT bFirstTime
THEN
	bDone := FALSE;                                 	(* Program done *)
	bBusy := FALSE;                                  	(* Program not busy *)
	bError := FALSE;                                 	(* Program not error *)
	udnErrorNo := 0;                                		(* Error number *)

	etLoadFromFile := ET_LoadFromFile_eWaitExecute;       				(* Next step *)
	
	bFirstTime := TRUE;
END_IF;

sPathName := CONCAT(
				sFilePath, CONCAT(
							sFileName, CONCAT(
										'.', sFileSuffix)));

rtExecute(CLK:= bExecute);				(* Positive edge for start *)

CASE etLoadFromFile OF
        
	ET_LoadFromFile_eWaitExecute:
		bBusy := FALSE;                                     		(* Program not busy *)
		bError := FALSE;                                    		(* Program not error *)

		IF rtExecute.Q
		THEN
			bDone := FALSE;                                 	(* Program done, in position *)
			bBusy := TRUE;                                  	(* Program busy *)
			udnErrorNo := 0;
			usnRowsCounter := 0;

			fbFileOpen.bExecute := FALSE;			(* File open *)
			fbFileClose.bExecute := FALSE;			(* File close *)
			fbFileGets.bExecute := FALSE;			(* File read *)

			dwMode := FOPEN_MODEREAD OR FOPEN_MODETEXT;

			etLoadFromFile := ET_LoadFromFile_eFileName;         		(* Next step *)
		END_IF;

	ET_LoadFromFile_eFileName:
		IF sFilePath <> ''
		     AND sFileName <> ''
		     AND sFileSuffix <> ''
		     AND byConfig <> 0
		THEN
			etLoadFromFile := ET_LoadFromFile_eChkFileExist;            			(* Next step *)

		ELSE
			udnErrorNo := ET_LoadFromFile_eFileName;

			etLoadFromFile := ET_LoadFromFile_eError;            			(* Next step *)

		END_IF

	ET_LoadFromFile_eChkFileExist:
		etLoadFromFile := ET_LoadFromFile_eFileOpen;            			(* Next step *)

	ET_LoadFromFile_eFileOpen:
		fbFileOpen.bExecute := TRUE;

		etLoadFromFile := ET_LoadFromFile_eChkFileOpen;            			(* Next step *)

	ET_LoadFromFile_eChkFileOpen:
		IF NOT fbFileOpen.bBusy
		     AND NOT fbFileOpen.bError
		THEN
			fbFileOpen.bExecute := FALSE;
			hFileHandle := fbFileOpen.hFile;

			MEMSET(ADR(arsData), 0, SIZEOF(arsData));						(* Array reset *)
			MEMSET(ADR(arbDataBool), 0, SIZEOF(arbDataBool));				(* Array reset *)
			MEMSET(ADR(arsDataDimRC), 0, SIZEOF(arsDataDimRC)); 		(* Array reset *)
			MEMSET(ADR(arrDataDimRC), 0, SIZEOF(arrDataDimRC)); 			(* Array reset *)

			etLoadFromFile := ET_LoadFromFile_eReadData;            			(* Next step *)

		ELSIF fbFileOpen.bError
		THEN
			fbFileOpen.bExecute := FALSE;
			udnErrorNo := fbFileOpen.nErrId;

			etLoadFromFile := ET_LoadFromFile_eError;            			(* Next step *)

		END_IF

	ET_LoadFromFile_eReadData:
		fbFileGets.bExecute := TRUE;

		etLoadFromFile := ET_LoadFromFile_eChkReadData;            			(* Next step *)

	ET_LoadFromFile_eChkReadData:
		IF NOT fbFileGets.bBusy
		     AND NOT fbFileGets.bError
		THEN
			fbFileGets.bExecute := FALSE;

			CASE byConfig OF
				1:	A_Option1();				(* Call option 1 *)
				2:	A_Option2();				(* Call option 2 *)
				3..4:	A_Option3();				(* Call option 3,4 *)
			END_CASE

		ELSIF fbFileGets.bError
		THEN
			fbFileGets.bExecute := FALSE;
			udnErrorNo := fbFileGets.nErrId;

			etLoadFromFile := ET_LoadFromFile_eError;            			(* Next step *)

		END_IF

	ET_LoadFromFile_eFileClose:
		fbFileClose.bExecute := TRUE;

		etLoadFromFile := ET_LoadFromFile_eChkFileClose;            			(* Next step *)

	ET_LoadFromFile_eChkFileClose:
		IF NOT fbFileClose.bBusy
		     AND NOT fbFileClose.bError
		THEN
			fbFileClose.bExecute := FALSE;

			IF NOT bError
			THEN
				etLoadFromFile := ET_LoadFromFile_eDone;            			(* Next step *)
			ELSE
				etLoadFromFile := ET_LoadFromFile_eError;            			(* Next step *)
			END_IF


		ELSIF fbFileClose.bError
		THEN
			fbFileClose.bExecute := FALSE;
			udnErrorNo := fbFileClose.nErrId;

			etLoadFromFile := ET_LoadFromFile_eError;            			(* Next step *)

		END_IF

	ET_LoadFromFile_eDone:
		bDone := TRUE;                                      		(* Program done, in position *)
		bBusy := FALSE;                                     		(* Program not busy *)
		bError := FALSE;
		udnErrorNo := 0;
	
		etLoadFromFile := ET_LoadFromFile_eNoExecute;            		(* Next step *)

	ET_LoadFromFile_eError:
		IF NOT bError
		     AND hFileHandle <> 0
		THEN
			bDone := FALSE;                                    	 	(* Program done, in position *)
			bError := TRUE;                                     		(* Program error *)
			bBusy := FALSE;                                     		(* Program not busy *)
	
			etLoadFromFile := ET_LoadFromFile_eFileClose;            		(* Next step *)

		ELSE
			bDone := FALSE;                                    	 	(* Program done, in position *)
			bError := TRUE;                                     		(* Program error *)
			bBusy := FALSE;                                     		(* Program not busy *)

			etLoadFromFile := ET_LoadFromFile_eNoExecute;            		(* Next step *)
		END_IF

	ET_LoadFromFile_eNoExecute:
		IF NOT bExecute
		THEN
			bDone := FALSE;                                 	(* Program done *)
			bBusy := FALSE;                                 	(* Program not busy *)
			bError := FALSE;                                		(* Program not error *)
			udnErrorNo := 0;
	
			etLoadFromFile := ET_LoadFromFile_eWaitExecute;       		(* Next step *)
	
		END_IF;
        
END_CASE;

fbFileOpen(
	sNetId := '',
	sPathName := sPathName,
	nMode := dwMode,
	ePath := PATH_GENERIC,
	tTimeout := tTimeout
);
fbFileClose(
	sNetId := '',
	hFile := hFileHandle,
	tTimeout := tTimeout
);

fbFileGets(
	sNetId := '',
	hFile :=  hFileHandle,
	tTimeout := tTimeout
);

ACTION A_Option1:
(* Option 1:

00000001 - 1 - Read line by line and save to array of string.

*)
(*****************************************************************************************************************************************************************************************************)

arsData[usnRowsCounter] := fbFileGets.sLine;											(* Read line (255 chars) from file *)

IF NOT fbFileGets.bEOF															(* Check received all data form file *)
THEN
	usnRowsCounter := usnRowsCounter + 1;
	etLoadFromFile := ET_LoadFromFile_eReadData;  									(* Read next line form file *)

ELSE
	etLoadFromFile := ET_LoadFromFile_eFileClose;  									(* Close current file *)

END_IF
END_ACTION

ACTION A_Option2:
(* Option 2:

00000010 - 2 - Read line by line. Save first signs to string and convert to array of bool.

*)
(*****************************************************************************************************************************************************************************************************)

sDataSign := fbFileGets.sLine;														(* Read first sign from line *)
sDataString := CONCAT(sDataString, sDataSign);										(* Created string of sign *)

ptString := ADR(sDataString);														(* Take adress to pointer of byte *)
arbyData :=  ptString^;																(* Take string into array of byte *)
arbDataBool[usnRowsCounter] := BYTE_TO_BOOL(arbyData[usnRowsCounter] AND 16#01);	(* Move data to Array of Bool *)

IF NOT fbFileGets.bEOF															(* Check received all data form file *)
THEN
	usnRowsCounter := usnRowsCounter + 1;
	etLoadFromFile := ET_LoadFromFile_eReadData;  									(* Read next line form file *)

ELSE
	etLoadFromFile := ET_LoadFromFile_eFileClose;  									(* Close current file *)

END_IF
END_ACTION

ACTION A_Option3:
(*Option 3:

00000011 - 3 - Transfer  array form file to array of string on PLC - requirements:
			- kind of columns separator (bySep) and sign end of line (byEndLine),
			- amount of rows (usiMaxDimR) and columns (usiMaxDimR) to read.

*)
(*****************************************************************************************************************************************************************************************************)

IF usnRowsCounter <= usnFileArrayMaxDimR 							(* Choose amount of rows from file *)
    AND NOT fbFileGets.bEOF
THEN
	arsData[usnRowsCounter] := fbFileGets.sLine; 						(* Read line (255 chars) from file *)

	ptByte := ADR(arsData[usnRowsCounter]);
	byDataSign :=  ptByte^;

	usnColumnsCounter := 0;
	REPEAT

		WHILE byDataSign <> F_ToASC(sSep) 			(* $T = HEX 09 *)   (* ; = HEX 3B *) (* EOF *)	(* Reaction for special sign in string*)
			      AND  byDataSign <> F_ToASC(sEndLine)	(* $N = HEX 0A *)
		DO
			IF byDataSign = F_ToASC(sComment)
			     OR byDataSign = F_ToASC('i')
			THEN
				EXIT;
			END_IF

			arsDataDimRC[usnRowsCounter , usnColumnsCounter] := CONCAT(arsDataDimRC[usnRowsCounter , usnColumnsCounter], F_ToCHR(byDataSign)); 	(* Read sign and create string*)

			IF byConfig = 4
			THEN
				IF F_CheckStringIsReal(arsDataDimRC[usnRowsCounter , usnColumnsCounter])
				THEN
					arrDataDimRC[usnRowsCounter , usnColumnsCounter] :=  STRING_TO_REAL(arsDataDimRC[usnRowsCounter , usnColumnsCounter]);				(* Create real *)
				ELSE
					udnErrorNo := 31;

					etLoadFromFile := ET_LoadFromFile_eError;            			(* Next step *)
					RETURN;
				END_IF
			END_IF

			ptByte := ptByte + 1;
			byDataSign :=  ptByte^;

		END_WHILE



		IF byDataSign <> F_ToASC(sEndLine)					(* Check end of line *)
		THEN
			IF byDataSign = F_ToASC(sComment)
			THEN
				EXIT;
			END_IF

			usnColumnsCounter := usnColumnsCounter + 1;			(* Set next columns *)
			ptByte := ptByte + 1;
			byDataSign :=  ptByte^;

		END_IF

	UNTIL byDataSign  = F_ToASC(sEndLine)					(* End when founds the end line sign*)
	END_REPEAT

	IF byDataSign <> F_ToASC(sComment)
	THEN
		usnRowsCounter := usnRowsCounter + 1;
	END_IF

	etLoadFromFile := ET_LoadFromFile_eReadData;  									(* Read next line form file *)

ELSE
	etLoadFromFile := ET_LoadFromFile_eFileClose;  									(* Close current file *)

END_IF
END_ACTION

END_FUNCTION_BLOCK

// ---- POUs/Tc2 Objects/String/F_CheckStringIsReal.TcPOU
FUNCTION F_CheckStringIsReal : BOOL (* TRUE if STR does not contain capital letters *)
VAR_INPUT
	str : T_MaxString;
END_VAR
VAR
	L : INT;
	pt : POINTER TO BYTE;
	pt2 : POINTER TO BYTE;
	pos: INT;
	pos2: INT;
END_VAR

pt := ADR(str);
pt2 := ADR(str);
L := LEN(str);

FOR pos := 1 TO L DO

	IF pt^ = 43 (* + *)
	     AND (pos <> 1)
	THEN
		F_CheckStringIsReal := FALSE;
		RETURN;

	ELSIF pt^ = 44 (* , *)
	THEN
		IF (pos = 1 (*OR pos = L*))
		THEN
			F_CheckStringIsReal := FALSE;
			RETURN;
		ELSE
			FOR pos2 := 1 TO L DO
				IF pos <> pos2
				THEN
					IF pt2^ = 44 OR pt2^ = 46
					THEN
						F_CheckStringIsReal := FALSE;
						RETURN;
					END_IF
				END_IF
				pt2 := pt2 + 1;
			END_FOR
		END_IF;
	ELSIF pt^ = 45 (* - *)
	     AND (pos <> 1)
	THEN
		F_CheckStringIsReal := FALSE;
		RETURN;
	ELSIF pt^ = 46 (* . *)
	THEN
		IF (pos = 1 (*OR pos = L*))
		THEN
			F_CheckStringIsReal := FALSE;
			RETURN;
		ELSE
			FOR pos2 := 1 TO L DO
				IF pos <> pos2
				THEN
					IF pt2^ = 44 OR pt2^ = 46
					THEN
						F_CheckStringIsReal := FALSE;
						RETURN;
					END_IF
				END_IF
				pt2 := pt2 + 1;
			END_FOR
		END_IF;
	ELSIF NOT (pt^ > 47 AND pt^ < 58)	(* 0 .. 9 *)
	     	    AND pt^ <> 43 (* + *)
	    	    AND pt^ <> 44 (* , *)
	             AND pt^ <> 45 (* - *)
	     	    AND pt^ <> 46 (* . *)
	THEN
		F_CheckStringIsReal := FALSE;
		RETURN;
	END_IF;

    	pt := pt + 1;
END_FOR;
F_CheckStringIsReal := L > 0;

END_FUNCTION

// ---- POUs/Machine/Group_0000 - General/Gr00Alarm/FB_Gr00Alarm.TcPOU
FUNCTION_BLOCK FB_Gr00Alarm
(*

The function block used to control general alarms of machine.

Constructor: 		Patryk Panylo
Company:		E. Riexinger GmbH
Date:			28.04.2015
Version:			1.00

Date:			Revision:		Who:				Comment
dd.mm.yyyy		x.xx			Initials			comment

*)
VAR_INPUT
	(* Input variables / Eingang Variablen *)
	etMachineMode				:ET_MachineMode;			(* Machine mode *)
	etMachineState				:ET_MachineState;			(* Machine state *)
	bNoEStop					:BOOL;						(* Emergency stop *)
	bConfirmAlarm				:BOOL;						(* Confirm alarm *)
	dtDateTime 					:DATE_AND_TIME;			(* Actual date and time *)
	nFatalErrorMaxIdx				:INT;						(* Maximal index of  using alarms *)
	nErrorMaxIdx					:INT;						(* Maximal index of  using alarms *)
	nWarningMaxIdx				:INT;						(* Maximal index of  using alarms *)
	nMessageMaxIdx				:INT;						(* Maximal index of  using alarms *)
	nHintMaxIdx					:INT;						(* Maximal index of  using alarms *)
	stAlarmIn						:ST_AlarmIn;					(* Alarm input *)
END_VAR
VAR_OUTPUT
	(* Output variables / Ausgang Variablen *)
	stAlarmOut					:ST_AlarmOut;				(* Alarm input *)
END_VAR
VAR_IN_OUT
	(* Input Output variables / Ausgang Variablen *)
	bMoveInterrupted				:BOOL;						(* Move interrupted *)
	bHomeCompleted				:BOOL;						(* Home completed *)
END_VAR
VAR
	(* Enummerations *)

	(* Variables *)

	(* References *)

	(* Interfaces *)

	(* Instances *)
	fbAlarm						:FB_Alarm;
END_VAR


(* Collection of alarms *)
fbAlarm(
	bEnable := TRUE,
	bNoEStop := bNoEStop,
	bReset := bConfirmAlarm,
	dtDateTime := dtDateTime,
	nFatalErrorMaxIdx := nFatalErrorMaxIdx,
	nErrorMaxIdx := nErrorMaxIdx,
	nWarningMaxIdx := nWarningMaxIdx,
	nMessageMaxIdx := nMessageMaxIdx,
	nHintMaxIdx := nHintMaxIdx,
    	stAlarmIn := stAlarmIn,
    	stAlarmOut => stAlarmOut
);

IF stAlarmOut.bFatalError
    OR stAlarmOut.bError
THEN
	(*bMoveInterrupted := FALSE;*)
	bHomeCompleted := FALSE;
END_IF;

END_FUNCTION_BLOCK

// ---- POUs/Tc2 Objects/Alarm/FB_Alarm.TcPOU
FUNCTION_BLOCK FB_Alarm
VAR_INPUT
	(* Input variables / Eingang Variablen *)
	bEnable					:BOOL;						(* Enable FB signal *)
	bNoEStop				:BOOL;						(* Emergency stop *)
	bReset					:BOOL;						(* Reset *)
	dtDateTime 				:DATE_AND_TIME;				(* Actual date and time *)
	nFatalErrorMaxIdx			:INT;						(* Maximal index of  using alarms *)
	nErrorMaxIdx				:INT;						(* Maximal index of  using alarms *)
	nWarningMaxIdx			:INT;						(* Maximal index of  using alarms *)
	nMessageMaxIdx			:INT;						(* Maximal index of  using alarms *)
	nHintMaxIdx				:INT;						(* Maximal index of  using alarms *)
	stAlarmIn					:ST_AlarmIn;					(* Alarm input *)
END_VAR
VAR_OUTPUT
	(* Output variables / Ausgang Variablen *)
	stAlarmOut				:ST_AlarmOut;				(* Alarm output *)
END_VAR
VAR
	(* Enummerations *)

	(* Variables *)
	arfbFatalError				:ARRAY[0..nALARM_MAX_NO] OF FB_FatalError;
	arfbError					:ARRAY[0..nALARM_MAX_NO] OF FB_Error;
	arfbWarning				:ARRAY[0..nALARM_MAX_NO] OF FB_Warning;
	arfbMessage				:ARRAY[0..nALARM_MAX_NO] OF FB_Message;
	arfbHint					:ARRAY[0..nALARM_MAX_NO] OF FB_Hint;

	nInc						:INT;

	(* References *)

	(* Interfaces *)

	(* Instances *)
	rtNoEStop				:R_TRIG;
	tonNoEStopDelay			:TON;
END_VAR

IF NOT bEnable
THEN
    RETURN;
END_IF;

IF dtDateTime = DT#1970-01-01-00:00
THEN
	RETURN;
END_IF

tonNoEStopDelay(
	IN := bNoEStop, 
	PT := T#1S
);
rtNoEStop(CLK := tonNoEStopDelay.Q);

stAlarmOut.bFatalError := FALSE;
stAlarmOut.bError := FALSE;
stAlarmOut.bWarning := FALSE;
stAlarmOut.bMessage := FALSE;
stAlarmOut.bHint := FALSE;

IF nFatalErrorMaxIdx > nALARM_MAX_NO
THEN
	nFatalErrorMaxIdx := nALARM_MAX_NO;
END_IF
FOR nInc := 0 TO nFatalErrorMaxIdx
DO
	(* ************************ FatalError ************************ *)
	stAlarmIn.arbFatalError[nInc].enType := ET_AlarmType_eFatalError;
	stAlarmIn.arbFatalError[nInc].dtDateTime := dtDateTime;
	
	arfbFatalError[nInc](
		bEnable := TRUE,
		stAlarmIn := stAlarmIn.arbFatalError[nInc]
	);

	stAlarmOut.arbFatalError[nInc].bActive := arfbFatalError[nInc].stAlarmOut.bActive;
	stAlarmOut.arbFatalError[nInc].dtDateTime := arfbFatalError[nInc].stAlarmOut.dtDateTime;
	stAlarmOut.arbFatalError[nInc].enType := arfbFatalError[nInc].stAlarmOut.enType;
	stAlarmOut.arbFatalError[nInc].dnCode := arfbFatalError[nInc].stAlarmOut.dnCode;
	
	stAlarmOut.bFatalError := stAlarmOut.bFatalError OR (stAlarmOut.arbFatalError[nInc].bActive > 0);
END_FOR

IF nErrorMaxIdx > nALARM_MAX_NO
THEN
	nErrorMaxIdx := nALARM_MAX_NO;
END_IF
FOR nInc := 0 TO nErrorMaxIdx
DO
	(* ************************ Error ************************ *)
	stAlarmIn.arbError[nInc].enType := ET_AlarmType_eError;
	stAlarmIn.arbError[nInc].dtDateTime := dtDateTime;
	
	arfbError[nInc](
		bEnable := TRUE,
		bReset := bReset OR rtNoEStop.Q,
		stAlarmIn := stAlarmIn.arbError[nInc]
	);

	stAlarmOut.arbError[nInc].bActive := arfbError[nInc].stAlarmOut.bActive;
	stAlarmOut.arbError[nInc].dtDateTime := arfbError[nInc].stAlarmOut.dtDateTime;
	stAlarmOut.arbError[nInc].enType := arfbError[nInc].stAlarmOut.enType;
	stAlarmOut.arbError[nInc].dnCode := arfbError[nInc].stAlarmOut.dnCode;
	
	stAlarmOut.bError := stAlarmOut.bError OR (stAlarmOut.arbError[nInc].bActive > 0);
END_FOR

IF nWarningMaxIdx > nALARM_MAX_NO
THEN
	nWarningMaxIdx := nALARM_MAX_NO;
END_IF
FOR nInc := 0 TO nWarningMaxIdx
DO
	(* ************************ Warning ************************ *)
	stAlarmIn.arbWarning[nInc].enType := ET_AlarmType_eWarning;
	stAlarmIn.arbWarning[nInc].dtDateTime := dtDateTime;
	
	arfbWarning[nInc](
		bEnable := TRUE,
		bReset := bReset OR rtNoEStop.Q,
		stAlarmIn := stAlarmIn.arbWarning[nInc]
	);
	
	stAlarmOut.arbWarning[nInc].bActive := arfbWarning[nInc].stAlarmOut.bActive;
	stAlarmOut.arbWarning[nInc].dtDateTime := arfbWarning[nInc].stAlarmOut.dtDateTime;
	stAlarmOut.arbWarning[nInc].enType := arfbWarning[nInc].stAlarmOut.enType;
	stAlarmOut.arbWarning[nInc].dnCode := arfbWarning[nInc].stAlarmOut.dnCode;
	
	stAlarmOut.bWarning := stAlarmOut.bWarning OR (stAlarmOut.arbWarning[nInc].bActive > 0);
END_FOR

IF nMessageMaxIdx > nALARM_MAX_NO
THEN
	nMessageMaxIdx := nALARM_MAX_NO;
END_IF
FOR nInc := 0 TO nMessageMaxIdx
DO
	(* ************************ Message ************************ *)
	stAlarmIn.arbMessage[nInc].enType := ET_AlarmType_eMessage;
	stAlarmIn.arbMessage[nInc].dtDateTime := dtDateTime;
	
	arfbMessage[nInc](
		bEnable := TRUE,
		stAlarmIn := stAlarmIn.arbMessage[nInc]
	);
	
	stAlarmOut.arbMessage[nInc].bActive := arfbMessage[nInc].stAlarmOut.bActive;
	stAlarmOut.arbMessage[nInc].dtDateTime := arfbMessage[nInc].stAlarmOut.dtDateTime;
	stAlarmOut.arbMessage[nInc].enType := arfbMessage[nInc].stAlarmOut.enType;
	stAlarmOut.arbMessage[nInc].dnCode := arfbMessage[nInc].stAlarmOut.dnCode;
		
	stAlarmOut.bMessage := stAlarmOut.bMessage OR (stAlarmOut.arbMessage[nInc].bActive > 0);
END_FOR

IF nHintMaxIdx > nALARM_MAX_NO
THEN
	nHintMaxIdx := nALARM_MAX_NO;
END_IF
FOR nInc := 0 TO nHintMaxIdx
DO
	(* ************************ Hint ************************ *)
	stAlarmIn.arbMessage[nInc].enType := ET_AlarmType_eMessage;
	stAlarmIn.arbMessage[nInc].dtDateTime := dtDateTime;
	
	arfbHint[nInc](
		bEnable := TRUE,
		stAlarmIn := stAlarmIn.arbHint[nInc]
	);

	stAlarmOut.arbHint[nInc].bActive := arfbHint[nInc].stAlarmOut.bActive;
	stAlarmOut.arbHint[nInc].dtDateTime := arfbHint[nInc].stAlarmOut.dtDateTime;
	stAlarmOut.arbHint[nInc].enType := arfbHint[nInc].stAlarmOut.enType;
	stAlarmOut.arbHint[nInc].dnCode := arfbHint[nInc].stAlarmOut.dnCode;
	
	stAlarmOut.bHint := stAlarmOut.bHint OR (stAlarmOut.arbHint[nInc].bActive > 0);
END_FOR

END_FUNCTION_BLOCK

// ---- POUs/Tc2 Objects/Alarm/FB_FatalError.TcPOU
FUNCTION_BLOCK FB_FatalError
VAR_INPUT
	(* Input variables / Eingang Variablen *)
	bEnable					:BOOL;						(* Enable FB signal *)
	stAlarmIn				:ST_AlarmProperties;				(* Alarm output *)
END_VAR
VAR_OUTPUT
	(* Output variables / Ausgang Variablen *)
	stAlarmOut				:ST_AlarmProperties;				(* Alarm output *)
END_VAR
VAR_IN_OUT

END_VAR
VAR
	(* Enummerations *)

	(* Variables *)

	(* References *)

	(* Interfaces *)

	(* Instances *)
	rtAlarm					:R_TRIG;
	ftAlarm					:F_TRIG;
END_VAR

(* Check method enabled *)
IF NOT bEnable
THEN
	RETURN;
END_IF;

rtAlarm(CLK := stAlarmIn.bActive);
ftAlarm(CLK := stAlarmIn.bActive);

IF rtAlarm.Q
THEN
	stAlarmOut.bActive := TRUE;
	stAlarmOut.enType := stAlarmIn.enType;
	stAlarmOut.dtDateTime := stAlarmIn.dtDateTime;
	stAlarmOut.dnCode := stAlarmIn.dnCode;
	
ELSIF ftAlarm.Q
THEN
	stAlarmOut.bActive := FALSE;
	(*stAlarmOut.enType := ET_AlarmType_eIdle;*)
	(*stAlarmOut.dtDateTime := DT#1970-01-01-00:00;*)
	(*stAlarmOut.dnCode := 0;*)
END_IF;

END_FUNCTION_BLOCK

// ---- POUs/Tc2 Objects/Alarm/FB_Error.TcPOU
FUNCTION_BLOCK FB_Error
VAR_INPUT
	(* Input variables / Eingang Variablen *)
	bEnable					:BOOL;						(* Enable FB signal *)
	bReset					:BOOL;						(* Reset *)
	stAlarmIn					:ST_AlarmProperties;			(* Alarm output *)
END_VAR
VAR_OUTPUT
	(* Output variables / Ausgang Variablen *)
	stAlarmOut				:ST_AlarmProperties;			(* Alarm output *)
END_VAR
VAR_IN_OUT

END_VAR
VAR
	(* Enummerations *)

	(* Variables *)

	(* References *)

	(* Interfaces *)

	(* Instances *)

END_VAR

(* Check method enabled *)
IF NOT bEnable
THEN
	RETURN;
END_IF;

IF bReset
THEN
	IF stAlarmOut.bActive
	THEN
		stAlarmOut.bActive := FALSE;
		(*stAlarmOut.enType := ET_AlarmType_eIdle;*)
		(*stAlarmOut.dtDateTime := DT#1970-01-01-00:00;*)
		(*stAlarmOut.dnCode := 0;*)
	END_IF;
ELSE
	IF stAlarmIn.bActive
	    AND NOT stAlarmOut.bActive
	THEN
		stAlarmOut.bActive := TRUE;
		stAlarmOut.enType := stAlarmIn.enType;
		stAlarmOut.dtDateTime := stAlarmIn.dtDateTime;
		stAlarmOut.dnCode := stAlarmIn.dnCode;
	END_IF;
END_IF;

END_FUNCTION_BLOCK

// ---- POUs/Tc2 Objects/Alarm/FB_Warning.TcPOU
FUNCTION_BLOCK FB_Warning
VAR_INPUT
	(* Input variables / Eingang Variablen *)
	bEnable					:BOOL;						(* Enable FB signal *)
	bReset					:BOOL;						(* Reset *)
	stAlarmIn					:ST_AlarmProperties;				(* Alarm output *)
END_VAR
VAR_OUTPUT
	(* Output variables / Ausgang Variablen *)
	bAlarmOut				:BOOL;				(* Alarm executed *)
	stAlarmOut				:ST_AlarmProperties;				(* Alarm output *)
END_VAR
VAR_IN_OUT

END_VAR
VAR
	(* Enummerations *)

	(* Variables *)

	(* References *)

	(* Interfaces *)

	(* Instances *)

END_VAR

(* Check method enabled *)
IF NOT bEnable
THEN
	RETURN;
END_IF;

IF bReset
THEN
	IF stAlarmOut.bActive
	THEN
		stAlarmOut.bActive := FALSE;
		(*stAlarmOut.enType := ET_AlarmType_eIdle;*)
		(*stAlarmOut.dtDateTime := DT#1970-01-01-00:00;*)
		(*stAlarmOut.dnCode := 0;*)
	END_IF;
	
ELSE
	IF stAlarmIn.bActive
	    AND NOT stAlarmOut.bActive
	THEN
		stAlarmOut.bActive := TRUE;
		stAlarmOut.enType := stAlarmIn.enType;
		stAlarmOut.dtDateTime := stAlarmIn.dtDateTime;
		stAlarmOut.dnCode := stAlarmIn.dnCode;
	END_IF;
	
END_IF;

END_FUNCTION_BLOCK

// ---- POUs/Tc2 Objects/Alarm/FB_Message.TcPOU
FUNCTION_BLOCK FB_Message
VAR_INPUT
	(* Input variables / Eingang Variablen *)
	bEnable					:BOOL;						(* Enable FB signal *)
	stAlarmIn				:ST_AlarmProperties;				(* Alarm output *)
END_VAR
VAR_OUTPUT
	(* Output variables / Ausgang Variablen *)
	stAlarmOut				:ST_AlarmProperties;				(* Alarm output *)
END_VAR
VAR_IN_OUT

END_VAR
VAR
	(* Enummerations *)

	(* Variables *)

	(* References *)

	(* Interfaces *)

	(* Instances *)
	rtAlarm					:R_TRIG;
	ftAlarm					:F_TRIG;
END_VAR

(* Check method enabled *)
IF NOT bEnable
THEN
	RETURN;
END_IF;

rtAlarm(CLK := stAlarmIn.bActive);
ftAlarm(CLK := stAlarmIn.bActive);

IF rtAlarm.Q
THEN
	stAlarmOut.bActive := TRUE;
	stAlarmOut.enType := stAlarmIn.enType;
	stAlarmOut.dtDateTime := stAlarmIn.dtDateTime;
	stAlarmOut.dnCode := stAlarmIn.dnCode;

ELSIF ftAlarm.Q
THEN
	stAlarmOut.bActive := FALSE;
	(*stAlarmOut.enType := ET_AlarmType_eIdle;*)
	(*stAlarmOut.dtDateTime := DT#1970-01-01-00:00;*)
	(*stAlarmOut.dnCode := 0;*)
END_IF;

END_FUNCTION_BLOCK

// ---- POUs/Tc2 Objects/Alarm/FB_Hint.TcPOU
FUNCTION_BLOCK FB_Hint
VAR_INPUT
	(* Input variables / Eingang Variablen *)
	bEnable					:BOOL;						(* Enable FB signal *)
	stAlarmIn					:ST_AlarmProperties;				(* Alarm output *)
END_VAR
VAR_OUTPUT
	(* Output variables / Ausgang Variablen *)
	stAlarmOut				:ST_AlarmProperties;				(* Alarm output *)
END_VAR
VAR_IN_OUT

END_VAR
VAR
	(* Enummerations *)

	(* Variables *)

	(* References *)

	(* Interfaces *)

	(* Instances *)
	rtAlarm					:R_TRIG;
	ftAlarm					:F_TRIG;
END_VAR

(* Check method enabled *)
IF NOT bEnable
THEN
	RETURN;
END_IF;

rtAlarm(CLK := stAlarmIn.bActive);
ftAlarm(CLK := stAlarmIn.bActive);

IF rtAlarm.Q
THEN
	stAlarmOut.bActive := TRUE;
	stAlarmOut.enType := stAlarmIn.enType;
	stAlarmOut.dtDateTime := stAlarmIn.dtDateTime;
	stAlarmOut.dnCode := stAlarmIn.dnCode;
    
ELSIF ftAlarm.Q
THEN
	stAlarmOut.bActive := FALSE;
	(*stAlarmOut.enType := ET_AlarmType_eIdle;*)
	(*stAlarmOut.dtDateTime := DT#1970-01-01-00:00;*)
	(*stAlarmOut.dnCode := 0;*)
END_IF;

END_FUNCTION_BLOCK

// ---- POUs/Machine/Group_0000 - General/Gr00Control/Gr00Safety/FB_Gr00Safety.TcPOU
FUNCTION_BLOCK FB_Gr00Safety
(*

The function block used to control genaeral safety of the machine.

Constructor: 		Patryk Panylo
Company:		E. Riexinger GmbH
Date:			28.04.2015
Version:			1.00

Date:			Revision:		Who:				Comment
dd.mm.yyyy		x.xx			Initials			comment

*)
VAR_INPUT
	(* Input variables / Eingang Variablen *)
	etMachineMode				:ET_MachineMode;			(* Machine mode *)
	etMachineState				:ET_MachineState;			(* Machine state *)
	bNoEStop					:BOOL;						(* No ermergency Stop / Keine Notaus *)
	bConfirmEStop				:BOOL;						(* Confirm no ermergency stop *)
	bMachineRunning				:BOOL;						(* Machine running / Maschine lauft *)
	arbPowerSupplyOn				:ARRAY [1..5] OF BOOL;		(* Power supply on / Leitung eingeschaltet *)
	bLightCurtain					:BOOL;						(* Light curtain ok / Freigabe Lichtschranke i.o *)
	bConfirmLightCurtain			:BOOL;						(* Confirm light Curtain input signal *)
	bAirPressure					:BOOL;						(* Air Pressure is available / Luftdruck ist vorhanden *)
	arbDoorsClosed				:ARRAY [1..5] OF BOOL;		(* Doors closed *)
	bDoorsClosed				:BOOL;						(* All doors closed *)
	bDoorsLocked				:BOOL;						(* All doors locked *)
	bDoorsLock					:BOOL;						(* All doors lock *)
	bTemperatur					:BOOL;						(* Temperatur *)
	stFieldbusStatus				:ST_FieldbusStatus;			(* Fieldbus status *)
	tFieldbusMasterStartUp		:TIME := T#30s;				(* Maximal start time for the fieldbus master *)
	tAirPressureOnDelay			:TIME := t#2s;					(* Delay air pressur on *)
	tAirPresentDelay				:TIME := t#2s;					(* Delay air pressur present *)
	tAirPressureBuildUp			:TIME := t#20s;				(* Max time to building up the air pressure  / Maximale Zeit zum erreichen des Solldrucks *)
	tLightCurtainDelay				:TIME := t#1s;					(* After time light Curtain safe *)
	tTempErrorDelay				:TIME := t#5m;					(* Max delay time until the message turns to an error *)
	tPowerSupplyOn				:TIME := t#2s;					(* Timeout power supply on *)
	tPowerSupplyOff				:TIME := t#1s;					(* Timeout power supply off *)
	tAdsTimeOut 					:TIME := t#2s;					(* Timout for ads commands / maximale zeit für die ausführung der ADS-Kommandos *)
END_VAR
VAR_OUTPUT
	(* Output variables / Ausgang Variablen *)
	bNoEmergencyStop			:BOOL;						(* No ermergency Stop / Keine Notaus *)
	bConfirmedEStop				:BOOL;						(* Confirmed emergency stop signal *)
	bFieldbusMasterOK			:BOOL;						(* Fieldbus master running *)
	bFieldbusBrake				:BOOL;						(* Fieldbus brake *)
	bAirPressureOK				:BOOL;						(* Air Pressure is available / Luftdruck ist vorhanden *)
	bAirPressureOn				:BOOL;						(* Air Pressure on / Luftdruck ein *)
	bPowerSupplyOk				:BOOL;						(* Power supply on / Leitung eingeschaltet *)
	bLightCurtainOK				:BOOL;						(* Light curtain ok / Freigabe Lichtschranke i.o *)
	bConfirmedLightCurtain			:BOOL;						(* Confirmed light Curtain signal *)
	bTemperaturOK				:BOOL;						(* Temperatur OK *)
	bAllDoorsLock				:BOOL;						(* All Doors lock / All Türen verriegeln *)
	bAllDoorsClosed				:BOOL;						(* All Doors closed / Alle Türen geschlossen *)
	bAllDoorsClosedLocked		:BOOL;						(* All Doors closed and locked / Alle Türen geschlossen und verrigelt *)
END_VAR
VAR_IN_OUT
	(* Input Output variables / Ausgang Variablen *)

END_VAR
VAR
	(* Enummerations *)

	(* Variables *)
	bFieldbusInit					:BOOL;						(* Fieldbus initialised *)

	(* References *)

	(* Interfaces *)

	(* Instances *)
	fbFieldbus					:FB_Fieldbus_v2;
	fbNoEmergencyStop			:FB_NoEmergencyStop;
	fbAirPressure					:FB_AirPressure;
	fbPowerSupply				:FB_PowerSupply;
	fbLightCurtain					:FB_LightCurtain;
	fbTemperatur					:FB_Temperature;
	fbDoorClosed				:ARRAY [1..5] OF FB_SignalWatchdog;

	tonFieldbusStartUp			:TON;
	fbFieldbusBreakWatchdog		:FB_SignalWatchdog;
END_VAR


A_Fieldbus();
A_EStop();
A_AirPressure();
A_PowerSupply();
A_LightCurtain();
A_Doors();
A_Temperatur();

ACTION A_AirPressure:

(* Air pressure controle *)
fbAirPressure(
	bEnable := TRUE,
	bIn := bAirPressure,
	bNoEStop := bNoEStop
			        AND bLightCurtainOK
			        AND bAllDoorsClosedLocked,
	tAirOnDelay := tAirPressureOnDelay,
	tAirPresentDelay := tAirPresentDelay,
	tTimeOut := tAirPressureBuildUp,
	bOut => bAirPressureOK,
	bAirOn => bAirPressureOn
);
END_ACTION

ACTION A_Doors:

(* Doors control *)
fbDoorClosed[1](
	bEnable := TRUE,
	bIn := arbDoorsClosed[1],
	tWatchdog := t#3s
);

bAllDoorsLock := bDoorsLock
			       OR bMachineRunning;
bAllDoorsClosed := bDoorsClosed;
bAllDoorsClosedLocked := bDoorsClosed
						AND bDoorsLocked;
END_ACTION

ACTION A_EStop:

(* Emergency stop controle *)
fbNoEmergencyStop(
	bEnable := TRUE,
	bIn := bNoEStop,
	bInConf := bConfirmEStop,
	bOut => bNoEmergencyStop,
	bOutConf => bConfirmedEStop
);
END_ACTION

ACTION A_Fieldbus:

(* Fieldbus controle *)
fbFieldbus(
	bEnable := TRUE,
	wFrmXWcState := stFieldbusStatus.wFrmXWcState,
	nMasterDeviceId := stFieldbusStatus.nMasterDeviceId,
	nMasterSlaveCount := stFieldbusStatus.nMasterSlaveCount,
	nMasterSlaveCountCfg := stFieldbusStatus.nMasterSlaveCountCfg,
	nMasterDevState := stFieldbusStatus.nMasterDevState,
	arrMasterNetId := stFieldbusStatus.arrMasterNetId,
	tTimeOut := tAdsTimeOut
);

IF fbFieldbus.bInit
    AND fbFieldbus.bDone
THEN
	IF fbFieldbus.bFieldbusOK
	     AND fbFieldbus.bFrameWcStateOK
	THEN
		bFieldbusInit := TRUE;
	END_IF;
END_IF

tonFieldbusStartUp(
	IN := NOT bFieldbusInit,
	PT := tFieldbusMasterStartUp
);

bFieldbusMasterOK := SEL(bFieldbusInit,
			   	        	        NOT tonFieldbusStartUp.Q,
			   	        	        NOT fbFieldbus.bMasterDevStateError);

bFieldbusBrake := bFieldbusInit
				AND NOT fbFieldbus.bMasterDevStateError
				AND (fbFieldbus.bFrameWcStateError
		  			  OR fbFieldbus.bSlaveCountError);
END_ACTION

ACTION A_LightCurtain:

(* Light Curtain control *)
fbLightCurtain(
	bEnable := TRUE,
	bIn := bLightCurtain,
	bInConf := bConfirmLightCurtain,
	tTimeOut := tLightCurtainDelay,
	bOut => bLightCurtainOK,
	bOutConf => bConfirmedLightCurtain
);
END_ACTION

ACTION A_PowerSupply:

(* Power supply control *)
fbPowerSupply(
	bEnable := TRUE,
	bIn := arbPowerSupplyOn[1]
		AND arbPowerSupplyOn[2]
		AND arbPowerSupplyOn[3]
		AND arbPowerSupplyOn[4]
		AND arbPowerSupplyOn[5],
	bNoEStop := bNoEStop,
	tPowerSupplyOn := tPowerSupplyOn,
	tPowerSupplyOff := tPowerSupplyOff,
	bOut => bPowerSupplyOk
);
END_ACTION

ACTION A_Temperatur:

fbTemperatur(
	bEnable := TRUE,
	bIn := bTemperatur,
	tTimeOut := tTempErrorDelay,
	bOut => bTemperaturOK,
 );
END_ACTION

END_FUNCTION_BLOCK

// ---- POUs/Tc2 Objects/Safety/Fieldbus/FB_Fieldbus_v2.TcPOU
FUNCTION_BLOCK FB_Fieldbus_v2
(*

The function block used to control fieldbus.

Constructor: 		Patryk Panylo
Company:		E. Riexinger GmbH
Date:			23.04.2015
Version:			1.00

Date:			Revision:		Who:				Comment
dd.mm.yyyy		x.xx			Initials			comment

*)
VAR_INPUT
	(* Input variables / Eingang Variablen *)
	bEnable					:BOOL;					(* Enable FB signal *)
	wFrmXWcState 			:WORD;					(* Link to task related ethercat frame state FrmXWcState *)
	nMasterDeviceId 			:UINT;
	nMasterSlaveCount		:UINT;
	nMasterSlaveCountCfg		:UINT;
	nMasterDevState			:UINT;
	arrMasterNetId			:T_AmsNetIdArr;
	tTimeOut					:TIME := t#5s;				(* Timeout for ADS commando *)
END_VAR
VAR_OUTPUT
	(* Output variables / Ausgang Variablen *)
	sMasterNetId				:T_AmsNetId ;			(* Fieldbus master ams net id*)
	bFieldbusOK				:BOOL;
	bFrameWcStateOK		:BOOL;
	bFrameWcStateError		:BOOL;
	bSlaveCountError			:BOOL;
	bMasterDevStateError		:BOOL;
	stMasterDevState			:ST_EcMasterDevState;
	bInit						:BOOL;
	bDone					:BOOL;					(* Program done *)
	bBusy					:BOOL;					(* Program busy  *)
	bError					:BOOL;					(* Program error  *)
	udnErrorNo				:UDINT;
	udnMessageNo			:UDINT;
	sMsg					:STRING;
END_VAR
VAR
	(* Enummerations *)

	(* Variables *)
	bFirstTime				:BOOL;
	wReqZeroMask			:WORD := 16#FFFF;		 (* Clear bit to ignore datagram error *)

	arstDiagSlaveInfo 			: ARRAY [0..dnDiagSlaveInfoMax] OF ST_SlaveStateInfo;
	arstDiagSlaveInfoScanned	: ARRAY [0..dnDiagSlaveInfoMax] OF ST_SlaveStateInfoScanned;

	(* References *)

	(* Interfaces *)

	(* Instances *)
	fbGetDeviceType			:IOF_GetDeviceType; 		(* Get the device type from the device ID *)
	fbEtherCATFrameDiag		:FB_EtherCATFrameDiag;
	fbEtherCATDiag			:FB_EtherCATDiag;
END_VAR
VAR CONSTANT
	dnDiagSlaveInfoMax			:DINT := 10;
END_VAR

IF NOT bEnable
THEN
	fbGetDeviceType(START := FALSE);
	bFieldbusOK := FALSE;
	bFrameWcStateOK := FALSE;
	bFrameWcStateError := FALSE;
	bSlaveCountError := FALSE;
	bMasterDevStateError := FALSE;
	bInit := FALSE;
	bDone := FALSE;
	bBusy := FALSE;
	bError := FALSE;
	udnErrorNo := 0;
	udnMessageNo := 0;
	sMsg := '';
	RETURN;
END_IF;


IF NOT bFirstTime
THEN
	bFieldbusOK := FALSE;
	bFrameWcStateOK := FALSE;
	bFrameWcStateError := FALSE;
	bSlaveCountError := FALSE;
	bMasterDevStateError := FALSE;
	bInit := FALSE;
	bDone := FALSE;
	bBusy := FALSE;
	bError := FALSE;
	udnErrorNo := 0;
	udnMessageNo := 0;
	sMsg := '';
	bFirstTime := TRUE;
END_IF;

(* Get the device type from the device ID *)
fbGetDeviceType(
	NETID := '',
	DEVICEID := nMasterDeviceId,
	START := TRUE,
	TMOUT := tTimeOut
);

(* Get the device type from the device ID *)
IF NOT fbGetDeviceType.BUSY 										(* No error *)
     AND NOT fbGetDeviceType.ERR
THEN

	CASE fbGetDeviceType.IODeviceType
	OF
		48: (* IODEVICETYPE_FC7500 	:= 48,  Beckhoff-SERCOS-PCI *)
			bInit := TRUE;
			bDone := FALSE;
			bBusy := FALSE;
			bError := FALSE;
			udnErrorNo := 0;											(* Error number *)
			(*bInitReady := unMasterState = 16#E005; 						(* Actual Phase is 4 *)
			bBreak := unMasterState = 16#E008;							(* Interrupt / Broke *)*)

		94: (* IODEVICETYPE_EtherCAT := 94,  Beckhoff-EtherCAT-PCI *)
			sMasterNetId := F_CreateAmsNetId(nIds := arrMasterNetId);
			bInit := sMasterNetID <> '' AND sMasterNetID <> '0.0.0.0.0.0';

			fbEtherCATFrameDiag(
				wFrmXWcState := wFrmXWcState,
				wReqZeroMask := wReqZeroMask,
				bFrameWcStateOK => bFrameWcStateOK
			);


			fbEtherCATDiag(
				sNetID := '',
				sMasterNetID	 := sMasterNetId,
				nMasterDevID := nMasterDeviceId,
				nSlaveCount := nMasterSlaveCount,
				nSlaveCountCfg := nMasterSlaveCountCfg,
				nMasterDevState := nMasterDevState,
				bAllFrameWcStatesOK	:= bFrameWcStateOK,
				tTimeout := tTimeOut,
				arstDiagSlaveInfo := arstDiagSlaveInfo,
				arstDiagSlaveInfoScanned	:= arstDiagSlaveInfoScanned,
				bEtherCATOK => bFieldbusOK,
				bFrameWcStateError	=> bFrameWcStateError,
				bSlaveCountError	=> bSlaveCountError,
				bMasterDevStateError=> bMasterDevStateError,
				stMasterDevState	=> stMasterDevState,
				bDone => bDone,
				bBusy => bBusy,
				bError => bError,
				iErrorID => udnErrorNo
			);

	ELSE (* IDLE *)
		bInit := FALSE;
		bDone := FALSE;
		bBusy := FALSE;
		bError := TRUE;
		udnErrorNo := 1;																			(* Error number *)
		sMsg := CONCAT('Unidentified fieldbus:', DINT_TO_STRING(fbGetDeviceType.IODeviceType));		(* Description error *)
	END_CASE;

ELSIF NOT fbGetDeviceType.BUSY
	    AND fbGetDeviceType.ERR
THEN
	bInit := FALSE;
	bDone := FALSE;
	bBusy := FALSE;
	bError := TRUE;
	udnErrorNo := 2;																				(* Error number *)
	sMsg := CONCAT('Fehler beim Lesen über ADS: ', UDINT_TO_STRING(fbGetDeviceType.ERRID));		(* Description error *)
	fbGetDeviceType(START := FALSE);
END_IF;

END_FUNCTION_BLOCK

// ---- POUs/Tc2 Objects/Safety/Fieldbus/FB_EtherCATFrameDiag.TcPOU
FUNCTION_BLOCK FB_EtherCATFrameDiag
VAR_INPUT
	wFrmXWcState 		: WORD;
	wReqZeroMask 		: WORD := 16#FFFF; (* bit TRUE: require wFrmXWcState.bit = FALSE, bit FALSE: ignore wFrmXWcState.bit *)
END_VAR
VAR_OUTPUT
	bFrameWcStateOK		: BOOL;
END_VAR
VAR
END_VAR

(* set/clear frame flag *)
bFrameWcStateOK := ((wFrmXWcState AND wReqZeroMask) = 0);

END_FUNCTION_BLOCK

// ---- POUs/Tc2 Objects/Safety/Fieldbus/FB_EtherCATDiag.TcPOU
FUNCTION_BLOCK FB_EtherCATDiag
(*

The function block used to control fieldbus.

Constructor: 		Patryk Panylo
Company:		E. Riexinger GmbH
Date:			22.11.2018
Version:			1.00

Date:			Revision:		Who:				Comment
dd.mm.yyyy		x.xx			Initials			comment

*)
VAR_INPUT
	(* Input variables / Eingang Variablen *)
	bEnable						:BOOL;						(* Enable FB signal *)
	sNetID						:T_AmsNetId; 				(* AmsNetId*)
	sMasterNetID					:T_AmsNetId; 				(* AmsNetId of the Fieldbus master device *)
	nMasterDevID				:UINT;
	nMasterDevState				:WORD;
	nSlaveCount 					:UINT;
	nSlaveCountCfg 				:UINT;
	bAllFrameWcStatesOK			:BOOL;
	tTimeout						:TIME := T#5s;
END_VAR
VAR_OUTPUT
	(* Output variables / Ausgang Variablen *)
	bDone						:BOOL;
	bBusy						:BOOL;
	bError						:BOOL;
	iErrorID						:UDINT;
	bEtherCATOK				:BOOL;
	bFrameWcStateError			:BOOL;
	bSlaveCountError				:BOOL;
	bMasterDevStateError			:BOOL;
	stMasterDevState				:ST_EcMasterDevState;
END_VAR
VAR_IN_OUT
	arstDiagSlaveInfo 				:ARRAY [0..dnDIAG_SLAVEINFO_SIZE] OF ST_SlaveStateInfo;
	arstDiagSlaveInfoScanned		:ARRAY [0..dnDIAG_SLAVEINFO_SIZE] OF ST_SlaveStateInfoScanned;
END_VAR
VAR
	(* Enummerations *)
	etEtherCATDiag				:ET_EtherCATDiag;

	(* Variables *)
	bFirstEtherCATOK				:BOOL;
	nMasterDevStatePrev			:WORD;
	bSlaveCountErrorPrev			:BOOL;
	bAllFrameWcStatesOKPrev		:BOOL;
	bDiagReq					:BOOL := TRUE;
	dnInc						:DINT;

	(* References *)

	(* Interfaces *)

	(* Instances *)


	(* -- Get Slave Addresses *)
	fbGetSlaveAddresses 			:FB_EcGetAllSlaveAddr;
	arrSlaveAddresses 			:ARRAY[0..iSLAVEADDR_ARR_SIZE] OF UINT;
	iNumOfSlavesRead			:INT;

	(* -- Get Slave States *)
	fbGetAllSlaveStates			:FB_EcGetAllSlaveStates;
	arrSlaveStates 				:ARRAY[0..iSLAVEADDR_ARR_SIZE] OF ST_EcSlaveState;

	(* -- Get Topology Data *)
	iTopologyData				:UDINT;
	fbGetTopologyData			:ADSREAD;
	arrTopologyData				:ARRAY[0..iSLAVEADDR_ARR_SIZE] OF ST_TopologyData;

	(* -- Check Topology *)
	iDiagIndex					:ARRAY [0..3] OF UINT;
	iDiagPort					:ARRAY [0..3] OF UINT;
	iIdx							:DINT;

	(* -- Scan Slaves *)
	fbEcGetScannedSlaves		:FB_EcGetScannedSlaves;
	arrScannedSlaveInfo			:ARRAY [0..iSLAVEADDR_ARR_SIZE] OF ST_EcSlaveScannedData;
	nScannedSlaves				:UINT;

	(* -- Get Slave Identities *)
	fbGetSlaveIdentity				:FB_EcGetSlaveIdentity;
	stIdentity 						:ST_EcSlaveIdentity;

	(* -- Get Slave Names *)
	fbGetSlaveName 				:IOF_GetBoxNameByAddr;
	strName						:STRING;

	arrSlaveInfo 					:ARRAY [0..iSLAVEADDR_ARR_SIZE] OF ST_SlaveStateInfo;
	arrSlaveInfoScanned			:ARRAY [0..iSLAVEADDR_ARR_SIZE] OF ST_SlaveStateInfoScanned;
END_VAR

(* cyclic diag *)
bFrameWcStateError := NOT bAllFrameWcStatesOK;

bSlaveCountError := (nSlaveCount <> nSlaveCountCfg) OR (nSlaveCount = 0);
IF (bSlaveCountError AND NOT bSlaveCountErrorPrev) OR (NOT bSlaveCountError AND bSlaveCountErrorPrev)
THEN
	bSlaveCountErrorPrev := bSlaveCountError;
	bDiagReq := TRUE;
END_IF

IF (bAllFrameWcStatesOK AND NOT bAllFrameWcStatesOKPrev) OR (NOT bAllFrameWcStatesOK AND bAllFrameWcStatesOKPrev)
THEN
	bAllFrameWcStatesOKPrev := bAllFrameWcStatesOK;
	bDiagReq := TRUE;
END_IF

IF (nMasterDevState <> nMasterDevStatePrev) THEN
	A_CheckMasterDevState();
	bDiagReq := TRUE;
END_IF

(* acyclic diag *)
CASE etEtherCATDiag OF

	ET_EtherCATDiag_eIdle:

		IF bDiagReq THEN
			bDiagReq := FALSE;

			IF sMasterNetID <> '' AND sMasterNetID <> '0.0.0.0.0.0'
			THEN
				bDone := FALSE;
				bBusy := TRUE;
				etEtherCATDiag := ET_EtherCATDiag_eGetSlaveAdresses;			(* Next step *)
			ELSE
				bError := TRUE;
				iErrorID := 7;
			END_IF

			bEtherCATOK := FALSE;
		ELSE
			IF (bSlaveCountError OR bMasterDevStateError OR NOT bAllFrameWcStatesOK) AND NOT (arrSlaveInfo[iDiagIndex[0]].bDiagData)
			THEN
				bEtherCATOK := FALSE;
				bDiagReq := TRUE;
			ELSIF (bSlaveCountError AND NOT bSlaveCountErrorPrev) OR (NOT bSlaveCountError AND bSlaveCountErrorPrev)
			THEN
				bSlaveCountErrorPrev := bSlaveCountError;
				bEtherCATOK := FALSE;
				bDiagReq := TRUE;
			ELSIF (nMasterDevState <> nMasterDevStatePrev)
			THEN
				bEtherCATOK := FALSE;
				bDiagReq := TRUE;
			ELSIF (bAllFrameWcStatesOK AND NOT bAllFrameWcStatesOKPrev) OR (NOT bAllFrameWcStatesOK AND bAllFrameWcStatesOKPrev)
			THEN
				bAllFrameWcStatesOKPrev := bAllFrameWcStatesOK;
				bEtherCATOK := FALSE;
				bDiagReq := TRUE;
			ELSIF (bSlaveCountError OR bMasterDevStateError OR NOT bAllFrameWcStatesOK OR arrSlaveInfo[iDiagIndex[0]].bDiagData)
			THEN
				bEtherCATOK := FALSE;
			ELSE
				bEtherCATOK := TRUE;
				IF NOT bFirstEtherCATOK
				THEN
					bFirstEtherCATOK := TRUE;
				END_IF
			END_IF
		END_IF

	ET_EtherCATDiag_eGetSlaveAdresses:
		A_GetSlaveAdresses();

	ET_EtherCATDiag_eGetSlaveStates:
		A_GetSlaveStates();

	ET_EtherCATDiag_eGetTopologyDataLen:
		A_GetTopoDataLen();

	ET_EtherCATDiag_eGetTopologyData:
		A_GetTopoData();

	ET_EtherCATDiag_eScanSlaves:
		A_ScanSlaves();

	ET_EtherCATDiag_eGetSlaveIdentity:
		A_GetSlaveIdentity();

	ET_EtherCATDiag_eGetSlaveName:
		A_GetSlaveName();

	ET_EtherCATDiag_eGetScannedSlaveName:
		A_GetScannedSlaveName();

	ET_EtherCATDiag_eDone:
		bDone := TRUE;
		bBusy := FALSE;
		etEtherCATDiag := ET_EtherCATDiag_eIdle;			(* Next step *)


END_CASE

ACTION A_CheckMasterDevState:
(* check master errors based on devstate *)
bMasterDevStateError := nMasterDevState <> 0;
stMasterDevState.bLinkError := ((nMasterDevState AND 16#000F) = 1) OR ((nMasterDevState AND 16#000F) = 4);
stMasterDevState.bResetRequired := ((nMasterDevState AND 16#000F) = 2) OR ((nMasterDevState AND 16#FFF0) = 16#10);
stMasterDevState.bMissFrmRedMode := (nMasterDevState AND 16#000F) = 8;
stMasterDevState.bWatchdogTriggerd := (nMasterDevState AND 16#20) = 16#20;
stMasterDevState.bDriverNotFound := (nMasterDevState AND 16#40) = 16#40;
stMasterDevState.bResetActive := (nMasterDevState AND 16#80) = 16#80;
stMasterDevState.bAtLeastOneNotInOp := ((nMasterDevState AND 16#100) = 16#100) OR ((nMasterDevState AND 16#200) = 16#200) OR
										((nMasterDevState AND 16#400) = 16#400) OR ((nMasterDevState AND 16#800) = 16#800);
stMasterDevState.bDcNotInSync := (nMasterDevState AND 16#1000) = 16#1000;
nMasterDevStatePrev := nMasterDevState;
END_ACTION

ACTION A_GetScannedSlaveName:
fbGetSlaveName(
	NETID := sNetID,
	DEVICEID := nMasterDevID,
	BOXADDR := arrScannedSlaveInfo[iDiagIndex[iIdx]].nAddr,
	START := TRUE,
	TMOUT := tTimeout,
	BOXNAME => strName
);

IF NOT fbGetSlaveName.BUSY
THEN
	fbGetSlaveName(START:= FALSE);

	(* add scanned info *)
	arrSlaveInfoScanned[iDiagIndex[iIdx]].nIndex 	:= iDiagIndex[iIdx] + 1;
	IF arrScannedSlaveInfo[iDiagIndex[iIdx]].nAddr <> 0
	THEN
		IF NOT fbGetSlaveName.ERR
		THEN
			arrSlaveInfoScanned[iDiagIndex[iIdx]].sName := strName;
		END_IF
	ELSE
		arrSlaveInfoScanned[iDiagIndex[iIdx]].sType := '';
	END_IF

	IF (iDiagIndex[iIdx] < nScannedSlaves)
	THEN
		arrSlaveInfoScanned[iDiagIndex[iIdx]].sType := F_ConvProductCodeToString(arrScannedSlaveInfo[iDiagIndex[iIdx]].stSlaveIdentity);
	ELSE
		arrSlaveInfoScanned[iDiagIndex[iIdx]].sType := '';
	END_IF

	arrSlaveInfoScanned[iDiagIndex[iIdx]].nECAddr := arrScannedSlaveInfo[iDiagIndex[iIdx]].nAddr;

	IF arrSlaveInfoScanned[iDiagIndex[iIdx]].sName <> arrSlaveInfo[iDiagIndex[iIdx]].sName
	THEN
		arrSlaveInfoScanned[iDiagIndex[iIdx]].bDifferentName := TRUE;
	ELSE
		arrSlaveInfoScanned[iDiagIndex[iIdx]].bDifferentName := FALSE;
	END_IF

	IF arrSlaveInfoScanned[iDiagIndex[iIdx]].nECAddr <> arrSlaveInfo[iDiagIndex[iIdx]].nECAddr
	THEN
		arrSlaveInfoScanned[iDiagIndex[iIdx]].bDifferentAddr := TRUE;
	ELSE
		arrSlaveInfoScanned[iDiagIndex[iIdx]].bDifferentAddr := FALSE;
	END_IF

	IF arrSlaveInfoScanned[iDiagIndex[iIdx]].sType <> arrSlaveInfo[iDiagIndex[iIdx]].sType
	THEN
		arrSlaveInfoScanned[iDiagIndex[iIdx]].bDifferentType := TRUE;
	ELSE
		arrSlaveInfoScanned[iDiagIndex[iIdx]].bDifferentType := FALSE;
	END_IF

	IF iIdx < 3
	THEN
		iIdx := iIdx + 1;

		etEtherCATDiag := ET_EtherCATDiag_eGetSlaveIdentity;			(* Next step *)
	ELSE
		iIdx := 0;

		FOR dnInc := 0 TO dnDIAG_SLAVEINFO_SIZE DO
			IF iDiagPort[dnInc] <> 0 THEN
				arstDiagSlaveInfo[dnInc] := arrSlaveInfo[iDiagIndex[dnInc]];
				arstDiagSlaveInfoScanned[dnInc] := arrSlaveInfoScanned[iDiagIndex[dnInc]];

				IF bFirstEtherCATOK
				THEN
					MEMSET(ADR(SaveDiagSlaveInfo[dnInc]), 0, SIZEOF(SaveDiagSlaveInfo[dnInc]));
					MEMSET(ADR(SaveDiagSlaveInfoScanned[dnInc]), 0, SIZEOF(SaveDiagSlaveInfoScanned[dnInc]));
					MEMCPY(ADR(SaveDiagSlaveInfo[dnInc]), ADR(arstDiagSlaveInfo[dnInc]), SIZEOF(arstDiagSlaveInfo[dnInc]));
					MEMCPY(ADR(SaveDiagSlaveInfoScanned[dnInc]), ADR(arstDiagSlaveInfoScanned[dnInc]), SIZEOF(arstDiagSlaveInfoScanned[dnInc]));
				END_IF
			ELSE
				MEMSET(ADR(arstDiagSlaveInfo[dnInc]), 0, SIZEOF(arstDiagSlaveInfo[dnInc]));
				MEMSET(ADR(arstDiagSlaveInfoScanned[dnInc]), 0, SIZEOF(arstDiagSlaveInfoScanned[dnInc]));
			END_IF
		END_FOR

		etEtherCATDiag := ET_EtherCATDiag_eDone;			(* Next step *)

	END_IF
END_IF
END_ACTION

ACTION A_GetSlaveAdresses:
fbGetSlaveAddresses(
	sNetId := sMasterNetID,
	pAddrBuf := ADR(arrSlaveAddresses),
	cbBufLen := SIZEOF(arrSlaveAddresses),
	bExecute := TRUE,
	tTimeout	:= tTimeout,
	nSlaves => iNumOfSlavesRead
);

IF NOT fbGetSlaveAddresses.bBusy
THEN
	fbGetSlaveAddresses(bExecute:= FALSE);

	IF NOT fbGetSlaveAddresses.bError
	THEN
		FOR dnInc := 0 TO MIN(iNumOfSlavesRead, iSLAVEADDR_ARR_SIZE)
		DO
			arrSlaveInfo[dnInc].nECAddr := arrSlaveAddresses[dnInc];
		END_FOR
	END_IF

	etEtherCATDiag := ET_EtherCATDiag_eGetSlaveStates;			(* Next step *)
END_IF
END_ACTION

ACTION A_GetSlaveIdentity:
fbGetSlaveIdentity(
	sNetId := sMasterNetID,
	nSlaveAddr := arrSlaveInfo[iDiagIndex[iIdx]].nECAddr,
	bExecute := TRUE,
	tTimeout	:= tTimeout,
	identity => stIdentity
);

IF NOT fbGetSlaveIdentity.bBusy
THEN
	fbGetSlaveIdentity(bExecute:= FALSE);

	IF NOT fbGetSlaveIdentity.bError
	THEN
		IF iDiagPort[iIdx] <> 0
		THEN
			arrSlaveInfo[iDiagIndex[iIdx]].nIndex	:= iDiagIndex[iIdx] + 1;
			arrSlaveInfo[iDiagIndex[iIdx]].sType 	:= F_ConvProductCodeToString(stSlaveIdentity := stIdentity);
		END_IF
	END_IF

	etEtherCATDiag := ET_EtherCATDiag_eGetSlaveName;			(* Next step *)
END_IF
END_ACTION

ACTION A_GetSlaveName:
fbGetSlaveName(
	NETID := sNetID,
	DEVICEID := nMasterDevID,
	BOXADDR := arrSlaveInfo[iDiagIndex[iIdx]].nECAddr,
	START := TRUE,
	TMOUT := tTimeout,
	BOXNAME => strName
);

IF NOT fbGetSlaveName.BUSY
THEN
	fbGetSlaveName(START:= FALSE);

	IF NOT fbGetSlaveName.ERR
	THEN
		IF iDiagPort[iIdx] <> 0
		THEN
			arrSlaveInfo[iDiagIndex[iIdx]].sName 	:= strName;
		END_IF
	END_IF

	etEtherCATDiag := ET_EtherCATDiag_eGetScannedSlaveName;			(* Next step *)
END_IF
END_ACTION

ACTION A_GetSlaveStates:
fbGetAllSlaveStates(
	sNetId := sMasterNetID,
	pStateBuf := ADR(arrSlaveStates),
	cbBufLen := SIZEOF(arrSlaveStates),
	bExecute := TRUE,
	tTimeout := tTimeout,
	nSlaves => iNumOfSlavesRead
);

IF NOT fbGetAllSlaveStates.bBusy
THEN
	fbGetAllSlaveStates(bExecute:= FALSE);

	IF NOT fbGetAllSlaveStates.bError
	THEN
		IF iNumOfSlavesRead = nSlaveCountCfg
		THEN
			FOR dnInc := 0 TO 3
			DO
				iDiagIndex[dnInc] := 0;
			END_FOR

			(* split slave state and link state *)
			FOR dnInc := 0 TO MIN(iNumOfSlavesRead, iSLAVEADDR_ARR_SIZE)
			DO
				(* slave state*)
				arrSlaveInfo[dnInc].stState.eEcState := arrSlaveStates[dnInc].deviceState AND 16#0F;
				arrSlaveInfo[dnInc].stState.bError := arrSlaveStates[dnInc].deviceState.4;
				arrSlaveInfo[dnInc].stState.bInvalidVPRS := arrSlaveStates[dnInc].deviceState.5;
				(* link state *)
				arrSlaveInfo[dnInc].stState.bNoCommToSlave := arrSlaveStates[dnInc].linkState.0;
				arrSlaveInfo[dnInc].stState.bLinkError := arrSlaveStates[dnInc].linkState.1;
				arrSlaveInfo[dnInc].stState.bMissingLink := arrSlaveStates[dnInc].linkState.2;
				arrSlaveInfo[dnInc].stState.bUnexpectedLink := arrSlaveStates[dnInc].linkState.3;
				arrSlaveInfo[dnInc].stState.bPortA := arrSlaveStates[dnInc].linkState.4;
				arrSlaveInfo[dnInc].stState.bPortB := arrSlaveStates[dnInc].linkState.5;
				arrSlaveInfo[dnInc].stState.bPortC := arrSlaveStates[dnInc].linkState.6;
				arrSlaveInfo[dnInc].stState.bPortD := arrSlaveStates[dnInc].linkState.7;
				(* DiagData *)
				arrSlaveInfo[dnInc].bDiagData := ((arrSlaveStates[dnInc].deviceState AND 16#F0) <> 0) OR
					(((arrSlaveStates[dnInc].deviceState AND 16#0F) > 0) AND ((arrSlaveStates[dnInc].deviceState AND 16#0F) < 8)) OR
					(arrSlaveStates[dnInc].linkState <> 0);

				IF arrSlaveInfo[dnInc].bDiagData
				THEN
					IF dnInc = 0
					THEN
						iDiagIndex[0] := 0;
					ELSE
						IF (iDiagIndex[0] = 0) AND NOT arrSlaveInfo[0].bDiagData
						THEN
							iDiagIndex[0] :=  DINT_TO_UINT(dnInc);
						END_IF
					END_IF
				END_IF
			END_FOR
		END_IF
	END_IF

	IF arrSlaveInfo[iDiagIndex[0]].bDiagData
	THEN
		etEtherCATDiag := ET_EtherCATDiag_eGetTopologyDataLen;			(* Next step *)
	ELSE
		FOR dnInc := 0 TO dnDIAG_SLAVEINFO_SIZE
		DO
			MEMSET(ADR(arstDiagSlaveInfo[dnInc]), 0, SIZEOF(arstDiagSlaveInfo[dnInc]));
			MEMSET(ADR(arstDiagSlaveInfoScanned[dnInc]), 0, SIZEOF(arstDiagSlaveInfoScanned[dnInc]));
		END_FOR

		etEtherCATDiag := ET_EtherCATDiag_eDone;			(* Next step *)
	END_IF
END_IF
END_ACTION

ACTION A_GetTopoData:
fbGetTopologyData(
	NETID := sMasterNetID,
	PORT := 16#FFFF,
	IDXGRP := 16#22,
	IDXOFFS := 0,
	LEN	 := iTopologyData * SIZEOF(arrTopologyData[0]),
	DESTADDR:= ADR(arrTopologyData),
	READ := TRUE,
	TMOUT := tTimeout,
);

IF NOT fbGetTopologyData.BUSY
THEN
	fbGetTopologyData(READ := FALSE);

	IF NOT fbGetTopologyData.ERR
	THEN
		iDiagPort[0] := arrTopologyData[iDiagIndex[0]].iOwnPhysicalAddr;
		iDiagPort[1] := arrTopologyData[iDiagIndex[0]].stPhysicalAddr.portB;
		iDiagPort[2] := arrTopologyData[iDiagIndex[0]].stPhysicalAddr.portC;
		iDiagPort[3] := arrTopologyData[iDiagIndex[0]].stPhysicalAddr.portD;

		(* clear diag index  *)
		iDiagIndex[1] := 0;
		iDiagIndex[2] := 0;
		iDiagIndex[3] := 0;

		(* find slaves on PortB of first slave with diag *)
		IF iDiagPort[1] <> 0
		THEN
			FOR dnInc := 0 TO MIN(iTopologyData-1,iSLAVEADDR_ARR_SIZE)
			DO
				IF arrTopologyData[dnInc].iOwnPhysicalAddr = iDiagPort[1]
				THEN
					iDiagIndex[1] :=  DINT_TO_UINT(dnInc);
					EXIT;
				END_IF
			END_FOR
		END_IF

		(* find slaves on PortC of first slave with diag *)
		IF iDiagPort[2] <> 0
		THEN
			FOR dnInc := 0 TO MIN(iTopologyData-1,iSLAVEADDR_ARR_SIZE)
			DO
				IF arrTopologyData[dnInc].iOwnPhysicalAddr = iDiagPort[2]
				THEN
					iDiagIndex[2] :=  DINT_TO_UINT(dnInc);
					EXIT;
				END_IF
			END_FOR
		END_IF

		(* find slaves on PortD of first slave with diag *)
		IF iDiagPort[3] <> 0
		THEN
			FOR dnInc := 0 TO MIN(iTopologyData-1,iSLAVEADDR_ARR_SIZE)
			DO
				IF arrTopologyData[dnInc].iOwnPhysicalAddr = iDiagPort[3]
				THEN
					iDiagIndex[3] :=  DINT_TO_UINT(dnInc);
					EXIT;
				END_IF
			END_FOR
		END_IF
	END_IF

	iIdx := 0;
	etEtherCATDiag := ET_EtherCATDiag_eScanSlaves;
END_IF
END_ACTION

ACTION A_GetTopoDataLen:
fbGetTopologyData(
	NETID := sMasterNetID,
	PORT := 16#FFFF,
	IDXGRP := EC_ADS_IGRP_MASTER_COUNT_SLAVE,
	IDXOFFS := EC_ADS_IOFFS_MASTER_COUNT_SLAVE,
	LEN	 := SIZEOF(iTopologyData),
	DESTADDR := ADR(iTopologyData),
	READ := TRUE,
	TMOUT := tTimeout,
);

IF NOT fbGetTopologyData.BUSY
THEN
	fbGetTopologyData(READ := FALSE);

	etEtherCATDiag := ET_EtherCATDiag_eGetTopologyData;			(* Next step *)
END_IF
END_ACTION

ACTION A_ScanSlaves:
fbEcGetScannedSlaves(
	bExecute := TRUE,
	sNetId := sMasterNetID,
	pArrEcScannedSlaveInfo := ADR(arrScannedSlaveInfo),
	cbBufLen := SIZEOF(arrScannedSlaveInfo),
	tTimeout := tTimeout
);

IF NOT fbEcGetScannedSlaves.bBusy
THEN
	fbEcGetScannedSlaves(bExecute := FALSE);

	IF fbEcGetScannedSlaves.bError THEN
		nScannedSlaves := 0;
	ELSE
		nScannedSlaves := fbEcGetScannedSlaves.nSlaves;
	END_IF

	etEtherCATDiag := ET_EtherCATDiag_eGetSlaveIdentity;
END_IF
END_ACTION

END_FUNCTION_BLOCK

// ---- POUs/Tc2 Objects/Safety/FB_NoEmergencyStop.TcPOU
FUNCTION_BLOCK FB_NoEmergencyStop
(*

The function block used to control emergency stop.

Constructor: 		Patryk Panylo
Company:		E. Riexinger GmbH
Date:			23.04.2015
Version:			1.00

Date:			Revision:		Who:				Comment
dd.mm.yyyy		x.xx			Initials			comment

*)
VAR_INPUT
	(* Input variables / Eingang Variablen *)
	bEnable					:BOOL;						(* Enable FB signal *)
	bIn						:BOOL;						(* Input signal *)
	bInConf					:BOOL;						(* Emergency stop *)
END_VAR
VAR_OUTPUT
	(* Output variables / Ausgang Variablen *)
	bOut					:BOOL;						(* Air pressure ok *)
	bOutConf					:BOOL;						(* Confirm output *)
	bError					:BOOL;						(* Error by no air pressure *)
	udnErrorNo				:UDINT;
	udnMessageNo			:UDINT;
	sMsg					:STRING;
END_VAR
VAR_IN_OUT

END_VAR
VAR
	(* Enummerations *)

	(* Variables *)
	bFirstTime				:BOOL;						(* First cycle *)

	(* References *)

	(* Interfaces *)

	(* Instances *)

END_VAR

IF NOT bEnable
THEN
	bOut := TRUE;
	bError := FALSE;
	udnErrorNo := 0;
	udnMessageNo := 0;
	sMsg := '';
	bFirstTime := FALSE;
	RETURN;
END_IF;

IF NOT bFirstTime
THEN
	bError := FALSE;
	udnErrorNo := 0;
	udnMessageNo := 0;
	sMsg := '';
	bFirstTime := TRUE;
END_IF;

bOut := bIn;
bError := NOT bOut;

IF bError
THEN
	udnErrorNo := 1;
	sMsg := 'Emergency stop';
ELSE
	udnErrorNo := 0;
	sMsg := 'No emergency stop';
END_IF;

bOutConf := bInConf AND NOT bIn;

END_FUNCTION_BLOCK

// ---- POUs/Tc2 Objects/Safety/FB_AirPressure.TcPOU
FUNCTION_BLOCK FB_AirPressure
(*

The function block used to control air pressure.

Constructor: 		Patryk Panylo
Company:		E. Riexinger GmbH
Date:			23.04.2015
Version:			1.00

Date:			Revision:		Who:				Comment
dd.mm.yyyy		x.xx			Initials			comment

*)
VAR_INPUT
	(* Input variables / Eingang Variablen *)
	bEnable					:BOOL;						(* Enable FB signal *)
	bIn						:BOOL;						(* Input signal *)
	bNoEStop				:BOOL;						(* Emergency stop *)
	tAirOnDelay				:TIME := t#2s;					(* Delay air pressure on *)
	tAirPresentDelay			:TIME := t#2s;					(* Delay air pressure present *)
	tTimeOut					:TIME := t#5s;					(* Timeout *)
END_VAR
VAR_OUTPUT
	(* Output variables / Ausgang Variablen *)
	bOut					:BOOL;						(* Air pressure ok *)
	bAirOn					:BOOL;						(* Air pressure on *)
	bError					:BOOL;						(* Error by no air pressure *)
	udnErrorNo				:UDINT;
	udnMessageNo			:UDINT;
	sMsg					:STRING;
END_VAR
VAR_IN_OUT

END_VAR
VAR
	(* Enummerations *)

	(* Variables *)
	bFirstTime				:BOOL;						(* First cycle *)

	(* References *)

	(* Interfaces *)

	(* Instances *)
	tonAirOnDelay			:TON;						(* Delay air pressure on *)
	tofAirPresentDelay		:TOF;						(* Delay air pressure present *)
	tonWatchDog				:TON;						(* Timer to delay *)
END_VAR

IF NOT bEnable
THEN
	bOut := TRUE;
	bError := FALSE;
	udnErrorNo := 0;
	udnMessageNo := 0;
	sMsg := '';
	tonWatchDog(IN := FALSE,
	             		 PT := tTimeOut);
	bFirstTime := FALSE;
	RETURN;
END_IF;

IF NOT bFirstTime
THEN
	bError := FALSE;
	udnErrorNo := 0;
	udnMessageNo := 0;
	sMsg := '';
	tonWatchDog(IN := FALSE,
	             		 PT := tTimeOut);
	bFirstTime := TRUE;
END_IF;

(* Air pressure on delay *)
tonAirOnDelay(
	IN := bNoEStop,
	PT := tAirOnDelay
);

bAirOn := tonAirOnDelay.Q;

(* Air pressure present delay *)
tofAirPresentDelay(
	IN := bIn,
	PT := tAirPresentDelay
);

bOut := tofAirPresentDelay.Q;

(* Timer starts when came rising edge of signal *)
tonWatchDog(
	IN := bAirOn,
	PT := tTimeOut
);

bError := NOT bOut
	        AND tonWatchDog.Q;

IF NOT bOut
     AND bAirOn
THEN
	IF tonWatchDog.Q                       		 (* Error if air pressure not present *)
	THEN
		udnErrorNo := 1;
		udnMessageNo := 0;
		sMsg := 'No pressured air';
	ELSE                                  				  (* Message if air pressure softstarting *)
		udnMessageNo := 1;
		sMsg := 'Air pressure building up';
	END_IF;
ELSE
	udnErrorNo := 0;
	udnMessageNo := 0;
	sMsg := '';
END_IF;

END_FUNCTION_BLOCK

// ---- POUs/Tc2 Objects/Safety/FB_PowerSupply.TcPOU
FUNCTION_BLOCK FB_PowerSupply
(*

The function block used to control power supply.

Constructor: 		Patryk Panylo
Company:		E. Riexinger GmbH
Date:			23.04.2015
Version:			1.00

Date:			Revision:		Who:				Comment
dd.mm.yyyy		x.xx			Initials			comment

*)
VAR_INPUT
	(* Input variables / Eingang Variablen *)
	bEnable					:BOOL;						(* Enable FB signal *)
	bIn						:BOOL;						(* Input signal *)
	bNoEStop				:BOOL;						(* Emergency stop *)
	tPowerSupplyOn			:TIME := t#2s;					(* Timeout power supply on *)
	tPowerSupplyOff			:TIME := t#1s;					(* Timeout power supply off *)
END_VAR
VAR_OUTPUT
	(* Output variables / Ausgang Variablen *)
	bOut					:BOOL;						(* Power supply ok *)
	bError					:BOOL;						(* Error by no air pressure *)
	udnErrorNo				:UDINT;
	udnMessageNo			:UDINT;
	sMsg					:STRING;
END_VAR
VAR_IN_OUT

END_VAR
VAR
	(* Enummerations *)

	(* Variables *)
	bFirstTime				:BOOL;						(* First cycle *)

	(* References *)

	(* Interfaces *)

	(* Instances *)
	tonPowerSupplyOn		:TON;						(* Timer to delay *)
	tofPowerSupplyOff			:TOF;						(* Timer to delay *)
END_VAR

IF NOT bEnable
THEN
	bOut := TRUE;
	bError := FALSE;
	udnErrorNo := 0;
	udnMessageNo := 0;
	sMsg := '';
	tonPowerSupplyOn(IN := FALSE,
				            PT := tPowerSupplyOn);
	tofPowerSupplyOff(IN := FALSE,
	            			 PT := tPowerSupplyOff);
	bFirstTime := FALSE;
    RETURN;
END_IF;

IF NOT bFirstTime
THEN
	bError := FALSE;
	udnErrorNo := 0;
	udnMessageNo := 0;
	sMsg := '';
	tonPowerSupplyOn(IN := FALSE,
	          			  PT := tPowerSupplyOn);
	tofPowerSupplyOff(IN := FALSE,
	             			 PT := tPowerSupplyOff);
	bFirstTime := TRUE;
END_IF;

(* Timer starts when came rising edge of signal *)
tonPowerSupplyOn(
	IN := bIn AND bNoEStop,
         PT := tPowerSupplyOn
);

tofPowerSupplyOff(
	IN := tonPowerSupplyOn.Q AND bNoEStop,
         PT := tPowerSupplyOff
);

bOut := tofPowerSupplyOff.Q;
bError := NOT tofPowerSupplyOff.Q;

IF bError
THEN
	udnErrorNo := 1;
	udnMessageNo := 0;
	sMsg := 'No power supply';
ELSE
	udnErrorNo := 0;
	udnMessageNo := 0;
	sMsg := '';
END_IF;

END_FUNCTION_BLOCK

// ---- POUs/Tc2 Objects/Safety/FB_LightCurtain.TcPOU
FUNCTION_BLOCK FB_LightCurtain
(*

The function block used to control light Curtain.

Constructor: 		Patryk Panylo
Company:		E. Riexinger GmbH
Date:			23.04.2015
Version:			1.00

Date:			Revision:		Who:				Comment
dd.mm.yyyy		x.xx			Initials			comment

*)
VAR_INPUT
	(* Input variables / Eingang Variablen *)
	bEnable					:BOOL;						(* Enable FB signal *)
	bIn						:BOOL;						(* Input signal *)
	bInConf					:BOOL;						(* Confirm *)
	tTimeOut					:TIME := t#1s;					(* Timeout *)
END_VAR
VAR_OUTPUT
	(* Output variables / Ausgang Variablen *)
	bOut					:BOOL;						(* Air pressure ok *)
	bOutConf					:BOOL;
	bError					:BOOL;						(* Error by no air pressure *)
	udnErrorNo				:UDINT;
	udnMessageNo			:UDINT;
	sMsg					:STRING;
END_VAR
VAR_IN_OUT

END_VAR
VAR
	(* Enummerations *)

	(* Variables *)
	bFirstTime				:BOOL;						(* First cycle *)

	(* References *)

	(* Interfaces *)

	(* Instances *)
	tonWatchDog				:TON;						(* Timer to delay *)
END_VAR

IF NOT bEnable
THEN
	bOut := TRUE;
	bError := FALSE;
	udnErrorNo := 0;
	udnMessageNo := 0;
	sMsg := '';
	tonWatchDog(IN := FALSE,
	             		 PT := tTimeOut);
	bFirstTime := FALSE;
	RETURN;
END_IF;

IF NOT bFirstTime
THEN
	bError := FALSE;
	udnErrorNo := 0;
	udnMessageNo := 0;
	sMsg := '';
	tonWatchDog(IN := FALSE,
				PT := tTimeOut);
	bFirstTime := TRUE;
END_IF;

(* Timer starts when came rising edge of signal *)
tonWatchDog(
	IN := bIn,
	PT := tTimeOut
);

bOut := tonWatchDog.Q;
bError := NOT bIn;

bOutConf := bInConf AND bError;

IF bError
THEN
	udnErrorNo := 1;
	sMsg := 'Light Curtain not ok';
    
ELSIF bOut
THEN
	udnErrorNo := 0;
	sMsg := 'Light curtain ok';
END_IF;

END_FUNCTION_BLOCK

// ---- POUs/Tc2 Objects/Safety/FB_Temperature.TcPOU
FUNCTION_BLOCK FB_Temperature
(*

The function block used to control temperature.

Constructor: 		Patryk Panylo
Company:		E. Riexinger GmbH
Date:			23.04.2015
Version:			1.00

Date:			Revision:		Who:				Comment
dd.mm.yyyy		x.xx			Initials			comment

*)
VAR_INPUT
	(* Input variables / Eingang Variablen *)
	bEnable					:BOOL;						(* Enable FB signal *)
	bIn						:BOOL;						(* Input signal *)
	tTimeOut					:TIME := t#5s;					(* Timeout *)
END_VAR
VAR_OUTPUT
	(* Output variables / Ausgang Variablen *)
	bOut					:BOOL;						(* Air pressure ok *)
	bError					:BOOL;						(* Error by no air pressure *)
	bWarning				:BOOL;						(* Warning by no temperature *)
	udnErrorNo				:UDINT;
	udnMessageNo			:UDINT;
	sMsg					:STRING;
END_VAR
VAR_IN_OUT

END_VAR
VAR
	(* Enummerations *)

	(* Variables *)
	bFirstTime				:BOOL;						(* First cycle *)

	(* References *)

	(* Interfaces *)

	(* Instances *)
	tonWatchDog				:TON;						(* Timer to delay *)
END_VAR

IF NOT bEnable
THEN
	bOut := TRUE;
	bError := FALSE;
	udnErrorNo := 0;
	udnMessageNo := 0;
	sMsg := '';
	tonWatchDog(IN := FALSE,
	             		 PT := tTimeOut);
	bFirstTime := FALSE;
	RETURN;
END_IF;

IF NOT bFirstTime
THEN
	bError := FALSE;
	udnErrorNo := 0;
	udnMessageNo := 0;
	sMsg := '';
	tonWatchDog(IN := FALSE,
	             		 PT := tTimeOut);
	bFirstTime := TRUE;
END_IF;

(* Timer starts when came rising edge of signal *)
tonWatchDog(
	IN := NOT bIn,
	PT := tTimeOut
);

bOut := bIn;
bError := NOT bOut
	        AND tonWatchDog.Q;
bWarning := NOT bError
		      AND NOT bOut;

IF NOT bOut
THEN
	IF tonWatchDog.Q                       		 (* Error if air pressure not present *)
	THEN
		udnErrorNo := 1;
		udnMessageNo := 0;
		sMsg := 'Temperature not ok';
	END_IF;
ELSE
	udnErrorNo := 0;
	udnMessageNo := 0;
	sMsg := '';
END_IF;

END_FUNCTION_BLOCK

